(* IEC 61131-3 sources: lasal-git-demo/CPU/LasalDemoProject/Class/_OpenSSL, 1 file *)

(* ---- _OpenSSL.st ---- *)
#include "..\..\Class\_OpenSSL\lsl_openssl.h"

(*!
<Class
	Name               = "_OpenSSL"
	Revision           = "1.9"
	RealtimeTask       = "false"
	CyclicTask         = "false"
	BackgroundTask     = "false"
	Sigmatek           = "true"
	OSInterface        = "true"
	HighPriority       = "false"
	Automatic          = "false"
	UpdateMode         = "Prescan"
	SharedCommandTable = "true"
	Objectsize         = "(284,120)"
	Comment            = "OpenSSL API">
	<Channels>
		<Server Name="ClassSvr" Visualized="false" Initialize="false" WriteProtected="true" Retentive="false"/>
	</Channels>
	<Dependencies>
		<Files>
			<File Path=".\Class\_OpenSSL\DefineCompiler.h" Include="false"/>
			<File Path=".\Class\_OpenSSL\lsl_c_openssl.h" Include="false"/>
			<File Path=".\Class\_OpenSSL\lsl_openssl.h" Include="true"/>
			<File Path=".\Source\code\OsiBaseNew.h" Include="false"/>
			<File Path=".\Source\code\OsiBaseNew.st"/>
		</Files>
	</Dependencies>
	<RevDoku>
		<Owner/>
		<Dokumentation Revision="1.9" Date="2022-09-02" Author="altman" Company="Sigmatek GmbH &amp; Co KG" Description="Fix function parameters for RSA_size and RSA_public_encrypt."/>
		<Dokumentation Revision="1.8" Date="2022-01-21" Author="altman" Company="Sigmatek GmbH &amp; Co KG" Description="The order of the function pointers (LSL_OPENSSL) has been corrected. &#13;&#10;Added new function (BIO_write, PEM_read_bio_RSA_PUBKEY, SHA512, SHA512_Init, SHA512_Update, SHA512_Final)&#13;&#10;Added new define NID_sha512"/>
		<Dokumentation Revision="1.7" Date="2020-05-05" Author="altman" Company="Sigmatek GmbH &amp; Co KG" Description="Added new function (EVP_sha256, SHA256)"/>
		<Dokumentation Revision="1.6" Date="2018-07-18" Author="FucHer" Company="Sigmatek GmbH &amp; Co KG" Description="Added comments for functions and parameters.&#13;&#10;d2i_RSAPrivateKey(): changed data type of parameter &lt;a&gt; from ^Void to ^pVoid.&#13;&#10;ASN1_TIME_set(): changed data type of parameter &lt;tx&gt; from ^DINT to DINT.&#13;&#10;Use dummy functions with a suitable return value."/>
		<Dokumentation Revision="1.5" Date="2018-06-19" Author="altman" Company="Sigmatek GmbH &amp; Co KG" Description="Added new function (X509_get_notBefore, X509_get_notAfter)&#13;&#10;Added new Type (ASN1_TIME)&#13;&#10;"/>
		<Dokumentation Revision="1.4" Date="2018-06-13" Author="altman" Company="Sigmatek GmbH &amp; Co KG" Description="Add new function (X509_cmp_time)&#13;&#10;Correct function parameter and CIL pointer name."/>
		<Dokumentation Revision="1.3" Date="2018-04-10" Author="altman" Company="Sigmatek GmbH &amp; Co KG" Description="Added new functions"/>
		<Dokumentation Revision="1.2" Date="2018-02-07" Author="fucher" Company="Sigmatek GmbH &amp; Co KG" Description="Added dummy functions to prevent fatal &quot;Ldr syntax error&quot; when CIL is not available.&#13;&#10;Removed duplicate entries from aMeths[]. Added missing entries to aMeths[].&#13;&#10;"/>
	</RevDoku>
</Class>
*)
_OpenSSL : CLASS
	TYPE
#pragma pack(push, 1)
	  LSL_OPENSSL : STRUCT
	    udVersion : UDINT;
	    udSize : UDINT;
	    d2i_X509 : pVoid;
	    X509_get_subject_name : pVoid;
	    X509_NAME_get_index_by_NID : pVoid;
	    X509_NAME_get_entry : pVoid;
	    X509_NAME_ENTRY_get_data : pVoid;
	    ASN1_STRING_to_UTF8 : pVoid;
	    OPENSSL_free : pVoid;
	    X509_free : pVoid;
	    SSLeay_version : pVoid;
	    OpenSSL_add_all_algorithms : pVoid;
	    ERR_load_crypto_strings : pVoid;
	    X509_STORE_CTX_get_ex_new_index : pVoid;
	    EVP_cleanup : pVoid;
	    CRYPTO_cleanup_all_ex_data : pVoid;
	    ERR_remove_state : pVoid;
	    ERR_free_strings : pVoid;
	    AES_set_encrypt_key : pVoid;
	    AES_set_decrypt_key : pVoid;
	    AES_cbc_encrypt : pVoid;
	    EVP_sha1 : pVoid;
	    HMAC : pVoid;
	    X509_STORE_free : pVoid;
	    X509_STORE_add_cert : pVoid;
	    SHA1 : pVoid;
	    RAND_bytes : pVoid;
	    RSA_generate_key : pVoid;
	    i2d_RSAPublicKey : pVoid;
	    i2d_RSAPrivateKey : pVoid;
	    d2i_RSAPrivateKey : pVoid;
	    d2i_PublicKey : pVoid;
	    d2i_PrivateKey : pVoid;
	    RSA_free : pVoid;
	    BIO_new_file : pVoid;
	    PEM_read_bio_PrivateKey : pVoid;
	    d2i_PKCS12_bio : pVoid;
	    PKCS12_parse : pVoid;
	    PKCS12_free : pVoid;
	    EVP_PKEY_get1_RSA : pVoid;
	    EVP_PKEY_free : pVoid;
	    BIO_free : pVoid;
	    PEM_write_bio_RSAPrivateKey : pVoid;
	    RSA_size : pVoid;
	    RSA_public_encrypt : pVoid;
	    RSA_private_decrypt : pVoid;
	    RSA_sign : pVoid;
	    ERR_get_error : pVoid;
	    ERR_error_string : pVoid;
	    RSA_verify : pVoid;
	    OBJ_txt2nid : pVoid;
	    X509_NAME_ENTRY_create_by_NID : pVoid;
	    X509_NAME_add_entry : pVoid;
	    X509V3_EXT_conf : pVoid;
	    X509_add_ext : pVoid;
	    X509_EXTENSION_free : pVoid;
	    X509_new : pVoid;
	    X509_set_version : pVoid;
	    X509_get_serialNumber : pVoid;
	    OPENSSL_Realloc : pVoid;
	    ASN1_INTEGER_set : pVoid;
	    X509_set_pubkey : pVoid;
	    X509_NAME_new : pVoid;
	    X509_set_subject_name : pVoid;
	    X509_set_issuer_name : pVoid;
	    X509_gmtime_adj : pVoid;
	    X509V3_set_ctx : pVoid;
	    X509_sign : pVoid;
	    X509_NAME_free : pVoid;
	    i2d_X509_bio : pVoid;
	    d2i_X509_bio : pVoid;
	    PEM_read_bio_X509 : pVoid;
	    X509_get_pubkey : pVoid;
	    OBJ_obj2nid : pVoid;
	    BIO_new : pVoid;
	    i2d_X509 : pVoid;
	    X509_verify : pVoid;
	    X509_STORE_new : pVoid;
	    CRYPTO_add_lock : pVoid;
	    X509_LOOKUP_file : pVoid;
	    X509_LOOKUP_ctrl : pVoid;
	    X509_verify_cert : pVoid;
	    X509_NAME_oneline : pVoid;
	    X509_load_crl_file : pVoid;
	    X509_STORE_CTX_new : pVoid;
	    X509_STORE_CTX_free : pVoid;
	    X509_STORE_CTX_init : pVoid;
	    X509_get_issuer_name : pVoid;
	    X509_LOOKUP_hash_dir : pVoid;
	    X509_STORE_set_flags : pVoid;
	    X509_STORE_add_lookup : pVoid;
	    X509_STORE_set_default_paths : pVoid;
	    X509_STORE_CTX_get_ex_data : pVoid;
	    X509_STORE_CTX_set_ex_data : pVoid;
	    X509_STORE_CTX_get_error : pVoid;
	    X509_STORE_CTX_get_current_cert : pVoid;
	    X509_STORE_CTX_get_error_depth : pVoid;
	    X509_verify_cert_error_string : pVoid;
	    i2d_PublicKey : pVoid;
	    EVP_PKEY_type : pVoid;
	    CRYPTO_realloc : pVoid;
	    BIO_ctrl : pVoid;
	    BIO_s_mem : pVoid;
	    BIO_s_file : pVoid;
	    X509_get_ext : pVoid;
	    EVP_PKEY_cmp : pVoid;
	    EVP_PKEY_new : pVoid;
	    ASN1_TIME_set : pVoid;
	    X509_CRL_sign : pVoid;
	    X509_PUBKEY_get : pVoid;
	    EVP_PKEY_assign : pVoid;
	    X509V3_EXT_print : pVoid;
	    X509_get_ext_by_NID : pVoid;
	    X509_CRL_set_version : pVoid;
	    X509_CRL_add0_revoked : pVoid;
	    X509_CRL_add1_ext_i2d : pVoid;
	    X509_CRL_set_lastUpdate : pVoid;
	    X509_CRL_set_nextUpdate : pVoid;
	    X509_NAME_add_entry_by_txt : pVoid;
	    X509_REVOKED_set_revocationDate : pVoid;
	    X509_CRL_set_issuer_name : pVoid;
	    X509_REVOKED_set_serialNumber : pVoid;
	    X509_NAME_ENTRY_free : pVoid;
	    X509_CRL_new : pVoid;
	    X509_CRL_free : pVoid;
	    ASN1_TIME_free : pVoid;
	    ASN1_INTEGER_new : pVoid;
	    ASN1_INTEGER_free : pVoid;
	    X509_REVOKED_new : pVoid;
	    X509_REVOKED_free : pVoid;
	    PEM_write_bio_X509_CRL : pVoid;
	    X509_cmp_time : pVoid;
	    X509_get_notBefore : pVoid;
	    X509_get_notAfter : pVoid;
	    EVP_sha256 : pVoid;
	    SHA256 : pVoid;
	    BIO_write : pVoid;
	    PEM_read_bio_RSA_PUBKEY : pVoid;
	    SHA512_Init : pVoid;
	    SHA512_Update : pVoid;
	    SHA512_Final : pVoid;
	    SHA512 : pVoid;
	  END_STRUCT;
#pragma pack(pop)
	END_TYPE
  //Servers:
	ClassSvr 	: SvrChCmd_DINT;
  //Clients:
  //Variables:
  //Functions:

	FUNCTION _OpenSSL
		VAR_OUTPUT
			ret_code 	: ConfStates;
		END_VAR;
				//! <Function Comment="Get the version of the OS interface." Name="GetVersion"/>
	FUNCTION VIRTUAL GLOBAL GetVersion
		VAR_OUTPUT
			ret0 	: UDINT;			//! <Variable Comment="&lt;&gt;0: version number of the OS interface&#13;&#10;  =0: error, no OpenSSL interface available." Name="GetVersion.ret0"/>
		END_VAR;
				//! <Function Comment="d2i_X509() attempts to decode &lt;len&gt; bytes at *&lt;in&gt;. If successful a pointer to the X509 structure is returned. If an error occurred, then NULL is returned.&#13;&#10;If &lt;px&gt; is not NULL, then the returned structure is written to *&lt;px&gt;. If *&lt;px&gt; is not NULL, then it is assumed that *&lt;px&gt; contains a valid X509 structure and an attempt is made to reuse it.&#13;&#10;This &quot;reuse&quot; capability is present for historical compatibility but its use is strongly discouraged (see BUGS in www.openssl.org/docs/man1.0.2/crypto/d2i_X509.html).&#13;&#10;&#13;&#10;NOTES&#13;&#10;The letters i and d in i2d_TYPE stand for &quot;internal&quot; (that is, an internal C structure) and &quot;DER&quot; respectively. So i2d_TYPE converts from internal to DER.&#13;&#10;&#13;&#10;If the call is successful *&lt;in&gt; is incremented to the byte following the parsed data.&#13;&#10;&#13;&#10;See also www.openssl.org/docs/man1.0.2/crypto/d2i_X509.html" Name="d2i_X509"/>
	FUNCTION __CDECL VIRTUAL GLOBAL d2i_X509
		VAR_INPUT
			px 	: ^pVoid;			//! <Variable Comment="Pointer to pointer to X509 structure (i.e. **X509).&#13;&#10;If &lt;px&gt; is not NULL, then the returned structure is written to *&lt;px&gt;." Name="d2i_X509.px"/>
			in 	: ^pChar;			//! <Variable Comment="Pointer to pointer to input buffer (i.e. **char)." Name="d2i_X509.in"/>
			len 	: DINT;			//! <Variable Comment="Number of bytes to decode." Name="d2i_X509.len"/>
		END_VAR
		VAR_OUTPUT
			RetAddr (EAX) 	: ^void;			//! <Variable Comment="If successful a pointer to the X509 structure is returned.&#13;&#10;If an error occurred, then NULL is returned. The error code that can be obtained by ERR_get_error()." Name="d2i_X509.RetAddr"/>
		END_VAR;
				//! <Function Comment="X509_get_subject_name() returns the subject name of certificate &lt;a&gt;. The returned value is an internal pointer which MUST NOT be freed.&#13;&#10;&#13;&#10;See also www.openssl.org/docs/man1.1.0/crypto/X509_get_subject_name.html" Name="X509_get_subject_name"/>
	FUNCTION __CDECL VIRTUAL GLOBAL X509_get_subject_name
		VAR_INPUT
			a 	: ^void;			//! <Variable Comment="Pointer to an X509 structure holding certificate &lt;a&gt;." Name="X509_get_subject_name.a"/>
		END_VAR
		VAR_OUTPUT
			RetAddr (EAX) 	: ^void;			//! <Variable Comment="RetAddr is a pointer to an X509_NAME structure.&#13;&#10;This pointer is an internal pointer which MUST NOT be freed." Name="X509_get_subject_name.RetAddr"/>
		END_VAR;
				//! <Function Comment="X509_NAME_get_index_by_NID() retrieves the next index matching &lt;nid&gt; after &lt;lastpos&gt;. &lt;lastpos&gt; should initially be set to -1.&#13;&#10;If there are no more entries -1 is returned. If &lt;nid&gt; is invalid (doesn&apos;t correspond to a valid OID) then -2 is returned.&#13;&#10;&#13;&#10;See also www.openssl.org/docs/man1.0.2/crypto/X509_NAME_get_entry.html" Name="X509_NAME_get_index_by_NID"/>
	FUNCTION __CDECL VIRTUAL GLOBAL X509_NAME_get_index_by_NID
		VAR_INPUT
			name 	: ^void;			//! <Variable Comment="Pointer to X509_NAME structure." Name="X509_NAME_get_index_by_NID.name"/>
			nid 	: DINT;			//! <Variable Comment="NID.&#13;&#10;Applications which could pass invalid NIDs to X509_NAME_get_index_by_NID() should check for the return value of -2." Name="X509_NAME_get_index_by_NID.nid"/>
			lastpos 	: DINT;			//! <Variable Comment="&lt;lastpos&gt; should initially be set to -1" Name="X509_NAME_get_index_by_NID.lastpos"/>
		END_VAR
		VAR_OUTPUT
			RetVal (EAX) 	: DINT;			//! <Variable Comment="Index of the next matching entry or -1 if not found.&#13;&#10;Method can also return -2 if the supplied NID is invalid." Name="X509_NAME_get_index_by_NID.RetVal"/>
		END_VAR;
				//! <Function Comment="X509_NAME_get_entry() retrieves the X509_NAME_ENTRY from &lt;name&gt; corresponding to index &lt;loc&gt;.&#13;&#10;Acceptable values for &lt;loc&gt; run from 0 to (X509_NAME_entry_count(&lt;name&gt;) - 1).&#13;&#10;The value returned is an internal pointer which must not be freed.&#13;&#10;&#13;&#10;See also www.openssl.org/docs/man1.0.2/crypto/X509_NAME_get_entry.html" Name="X509_NAME_get_entry"/>
	FUNCTION __CDECL VIRTUAL GLOBAL X509_NAME_get_entry
		VAR_INPUT
			name 	: ^void;			//! <Variable Comment="Pointer to X509_NAME structure." Name="X509_NAME_get_entry.name"/>
			loc 	: DINT;			//! <Variable Comment="0 to (X509_NAME_entry_count(name) - 1)" Name="X509_NAME_get_entry.loc"/>
		END_VAR
		VAR_OUTPUT
			RetAddr (EAX) 	: ^void;			//! <Variable Comment="Pointer to an X509_NAME_ENTRY structure.&#13;&#10;This is an internal pointer which MUST NOT be freed." Name="X509_NAME_get_entry.RetAddr"/>
		END_VAR;
				//! <Function Comment="X509_NAME_ENTRY_get_data() retrieves the field value of &lt;NeAddr&gt; in an ASN1_STRING structure.&#13;&#10;&#13;&#10;See also www.openssl.org/docs/man1.1.0/crypto/X509_NAME_ENTRY_get_data.html" Name="X509_NAME_ENTRY_get_data"/>
	FUNCTION __CDECL VIRTUAL GLOBAL X509_NAME_ENTRY_get_data
		VAR_INPUT
			NeAddr 	: ^void;			//! <Variable Comment="Pointer to X509_NAME_ENTRY structure." Name="X509_NAME_ENTRY_get_data.NeAddr"/>
		END_VAR
		VAR_OUTPUT
			RetAddr (EAX) 	: ^void;			//! <Variable Comment="Pointer to ASN1_STRING structure." Name="X509_NAME_ENTRY_get_data.RetAddr"/>
		END_VAR;
				//! <Function Comment="ASN1_STRING_to_UTF8() converts the string &lt;in&gt; to UTF8 format, the converted data is allocated in a buffer in *&lt;out&gt;.&#13;&#10;The length of &lt;out&gt; is returned or a negative error code. The buffer *&lt;out&gt; should be freed using OPENSSL_free().&#13;&#10;&#13;&#10;See also www.openssl.org/docs/man1.1.0/crypto/ASN1_STRING_to_UTF8.html" Name="ASN1_STRING_to_UTF8"/>
	FUNCTION __CDECL VIRTUAL GLOBAL ASN1_STRING_to_UTF8
		VAR_INPUT
			out 	: ^pChar;			//! <Variable Comment="Pointer to pointer to output buffer (i.e. **char)." Name="ASN1_STRING_to_UTF8.out"/>
			in 	: ^void;			//! <Variable Comment="Pointer to ASN1_STRING structure." Name="ASN1_STRING_to_UTF8.in"/>
		END_VAR
		VAR_OUTPUT
			RetVal (EAX) 	: DINT;			//! <Variable Comment="The length of &lt;out&gt; or a negative error code." Name="ASN1_STRING_to_UTF8.RetVal"/>
		END_VAR;
				//! <Function Comment="OPENSSL_free() is like the C free() function.&#13;&#10;&#13;&#10;See also www.openssl.org/docs/man1.1.0/crypto/OPENSSL_malloc.html" Name="OPENSSL_free"/>
	FUNCTION __CDECL VIRTUAL GLOBAL OPENSSL_free
		VAR_INPUT
			Addr 	: ^void;			//! <Variable Comment="Void pointer to the buffer that should be freed." Name="OPENSSL_free.Addr"/>
		END_VAR;
				//! <Function Comment="X509_free() frees up the X509 structure &lt;a&gt;.&#13;&#10;&#13;&#10;See also www.openssl.org/docs/man1.0.2/crypto/X509_free.html" Name="X509_free"/>
	FUNCTION __CDECL VIRTUAL GLOBAL X509_free
		VAR_INPUT
			a 	: ^void;			//! <Variable Comment="Pointer to an X509 structure." Name="X509_free.a"/>
		END_VAR;
				//! <Function Comment="SSLeay_version() returns a pointer to a constant string describing the version of the OpenSSL library or giving information about the library build.&#13;&#10;&#13;&#10;See also www.openssl.org/docs/man1.0.2/crypto/SSLeay_version.html" Name="SSLeay_version"/>
	FUNCTION __CDECL VIRTUAL GLOBAL SSLeay_version
		VAR_INPUT
			info_type 	: DINT;			//! <Variable Comment="The following values are supported:&#13;&#10;&#13;&#10;SSLEAY_VERSION&#13;&#10;  The version of the OpenSSL library including the release date.&#13;&#10;SSLEAY_CFLAGS&#13;&#10;  The compiler flags set for the compilation process in the form &quot;compiler: ...&quot; if available or &quot;compiler: information not available&quot; otherwise.&#13;&#10;SSLEAY_BUILT_ON&#13;&#10;  The date of the build process in the form &quot;built on: ...&quot; if available or &quot;built on: date not available&quot; otherwise.&#13;&#10;SSLEAY_PLATFORM&#13;&#10;  The &quot;Configure&quot; target of the library build in the form &quot;platform: ...&quot; if available or &quot;platform: information not available&quot; otherwise.&#13;&#10;SSLEAY_DIR&#13;&#10;  The &quot;OPENSSLDIR&quot; setting of the library build in the form &quot;OPENSSLDIR: &quot;...&quot; if available or &quot;OPENSSLDIR: N/A&quot; otherwise.&#13;&#10;" Name="SSLeay_version.info_type"/>
		END_VAR
		VAR_OUTPUT
			RetAddr (EAX) 	: ^CHAR;			//! <Variable Comment="The following return values can occur:&#13;&#10;&quot;not available&quot;&#13;&#10;  An invalid value for info_type was given.&#13;&#10;Pointer to constant string&#13;&#10;  Textual description.&#13;&#10;" Name="SSLeay_version.RetAddr"/>
		END_VAR;
				//! <Function Comment="OpenSSL keeps an internal table of digest algorithms and ciphers. It uses this table to lookup ciphers via functions such as EVP_get_cipher_byname().&#13;&#10;OpenSSL_add_all_algorithms() adds all algorithms (digests and ciphers) to the table.&#13;&#10;&#13;&#10;See also www.openssl.org/docs/man1.1.0/crypto/OpenSSL_add_all_algorithms.html&#13;&#10;and       https://wiki.openssl.org/index.php/Libcrypto_API" Name="OpenSSL_add_all_algorithms"/>
	FUNCTION __CDECL VIRTUAL GLOBAL OpenSSL_add_all_algorithms;
				//! <Function Comment="ERR_load_crypto_strings() registers the error strings for all libcrypto functions.&#13;&#10;This function should be called before generating textual error messages. However, this is not required when memory usage is an issue.&#13;&#10;&#13;&#10;See also www.openssl.org/docs/man1.0.2/crypto/ERR_load_crypto_strings.html&#13;&#10;and       https://wiki.openssl.org/index.php/Libcrypto_API" Name="ERR_load_crypto_strings"/>
	FUNCTION __CDECL VIRTUAL GLOBAL ERR_load_crypto_strings;
				//! <Function Comment="The X509_STORE_CTX_get_ex_new_index() function is initially called to &quot;register&quot; some new application specific data.&#13;&#10;It takes three optional function pointers which are called when the parent structure (in this case an RSA structure) is initially created, when it is copied and when it is freed up.&#13;&#10;If any or all of these function pointer arguments are not used they should be set to NULL.&#13;&#10;It also takes additional long and pointer parameters which will be passed to the supplied functions new_func(), dup_func() and free_func() but which otherwise have no special meaning.&#13;&#10;&#13;&#10;See also www.openssl.org/docs/man1.0.2/crypto/X509_STORE_CTX_get_ex_new_index.html&#13;&#10;and       www.openssl.org/docs/man1.0.2/crypto/RSA_get_ex_new_index.html" Name="X509_STORE_CTX_get_ex_new_index"/>
	FUNCTION __CDECL VIRTUAL GLOBAL X509_STORE_CTX_get_ex_new_index
		VAR_INPUT
			argl 	: DINT;			//! <Variable Comment="Will be passed to the supplied functions &lt;new_func&gt;, &lt;dup_func&gt;, &lt;free_func&gt;." Name="X509_STORE_CTX_get_ex_new_index.argl"/>
			argp 	: ^void;			//! <Variable Comment="Will be passed to the supplied functions &lt;new_func&gt;, &lt;dup_func&gt;, &lt;free_func&gt;." Name="X509_STORE_CTX_get_ex_new_index.argp"/>
			new_func 	: ^void;			//! <Variable Comment="Optional function pointer CRYPTO_EX_new which is called when the parent structure (in this case an RSA structure) is initially created.&#13;&#10;&#13;&#10;typedef int CRYPTO_EX_new(void *parent, void *ptr, CRYPTO_EX_DATA *ad, int idx, long argl, void *argp);" Name="X509_STORE_CTX_get_ex_new_index.new_func"/>
			dup_func 	: ^void;			//! <Variable Comment="Optional function pointer CRYPTO_EX_dup which is called when the parent structure (in this case an RSA structure) is copied.&#13;&#10;&#13;&#10;typedef int CRYPTO_EX_dup(CRYPTO_EX_DATA *to, CRYPTO_EX_DATA *from, void *from_d, int idx, long argl, void *argp);" Name="X509_STORE_CTX_get_ex_new_index.dup_func"/>
			free_func 	: ^void;			//! <Variable Comment="Optional function pointer CRYPTO_EX_free which is called when the parent structure (in this case an RSA structure) is freed up.&#13;&#10;&#13;&#10;typedef void CRYPTO_EX_free(void *parent, void *ptr, CRYPTO_EX_DATA *ad, int idx, long argl, void *argp);" Name="X509_STORE_CTX_get_ex_new_index.free_func"/>
		END_VAR
		VAR_OUTPUT
			RetVal (EAX) 	: DINT;			//! <Variable Comment="Returns a new index or -1 on failure (note 0 is a valid index value).&#13;&#10;Each successful call will return an index greater than any previously returned." Name="X509_STORE_CTX_get_ex_new_index.RetVal"/>
		END_VAR;
				//! <Function Comment="EVP_cleanup() removes all ciphers and digests from the table used by OpenSSL_add_all_algorithms().&#13;&#10;&#13;&#10;See also www.openssl.org/docs/man1.0.2/crypto/OpenSSL_add_all_algorithms.html&#13;&#10;and       https://wiki.openssl.org/index.php/Libcrypto_API" Name="EVP_cleanup"/>
	FUNCTION __CDECL VIRTUAL GLOBAL EVP_cleanup;
				//! <Function Comment="OpenSSL provides two primary libraries: libssl and libcrypto. The libcrypto library provides the fundamental cryptographic routines used by libssl. &#13;&#10;You can however use libcrypto without using libssl. In order to use libcrypto it must first be initialised.&#13;&#10;Call EVP_cleanup() and CRYPTO_cleanup_all_ex_data() do to the necessary cleanup after using the libcrypto routines.&#13;&#10;&#13;&#10;See also https://wiki.openssl.org/index.php/Libcrypto_API" Name="CRYPTO_cleanup_all_ex_data"/>
	FUNCTION __CDECL VIRTUAL GLOBAL CRYPTO_cleanup_all_ex_data;
				//! <Function Comment="ERR_remove_state() frees the error queue associated with the current thread.&#13;&#10;Since threads in OpenSSL are no longer identified by unsigned long values any argument to this function is ignored.&#13;&#10;&#13;&#10;Since error queue data structures are allocated automatically for new threads, they must be freed when threads are terminated in order to avoid memory leaks.&#13;&#10;&#13;&#10;See also www.openssl.org/docs/man1.0.2/crypto/ERR_remove_state.html" Name="ERR_remove_state"/>
	FUNCTION __CDECL VIRTUAL GLOBAL ERR_remove_state
		VAR_INPUT
			pid 	: UDINT;			//! <Variable Comment="Since threads in OpenSSL are no longer identified by unsigned long values any argument to this function is ignored." Name="ERR_remove_state.pid"/>
		END_VAR;
				//! <Function Comment="ERR_free_strings() frees all previously loaded error strings.&#13;&#10;&#13;&#10;See also www.openssl.org/docs/man1.0.2/crypto/ERR_free_strings.html" Name="ERR_free_strings"/>
	FUNCTION __CDECL VIRTUAL GLOBAL ERR_free_strings;
				//! <Function Comment="AES_set_encrypt_key() configures &lt;key&gt; to encrypt with the &lt;bits&gt;-bit key, &lt;userkey&gt;.&#13;&#10;&#13;&#10;&lt;userkey&gt; contains the actual 128-bit AES key. &lt;key&gt; is a data structure holding a transformed version of the &lt;userkey&gt;, for efficiency.&#13;&#10;&#13;&#10;See also https://boringssl.googlesource.com/boringssl/+/2490/include/openssl/aes.h&#13;&#10;and       www.cs.umd.edu/~jkatz/security/example.c" Name="AES_set_encrypt_key"/>
	FUNCTION __CDECL VIRTUAL GLOBAL AES_set_encrypt_key
		VAR_INPUT
			userkey 	: ^USINT;			//! <Variable Comment="Pointer to actual 128-bit AES key." Name="AES_set_encrypt_key.userkey"/>
			bits 	: DINT;			//! <Variable Comment="Number of bits in &lt;userkey&gt;." Name="AES_set_encrypt_key.bits"/>
			key 	: ^void;			//! <Variable Comment="Pointer to an AES_KEY structure. It holds a transformed version of the &lt;userkey&gt;, for efficiency." Name="AES_set_encrypt_key.key"/>
		END_VAR
		VAR_OUTPUT
			RetVal (EAX) 	: DINT;			//! <Variable Comment="WARNING: unlike other OpenSSL functions, this returns zero on success and a negative number on error." Name="AES_set_encrypt_key.RetVal"/>
		END_VAR;
				//! <Function Comment="AES_set_decrypt_key() configures &lt;key&gt; to decrypt with the &lt;bits&gt;-bit key, &lt;userkey&gt;.&#13;&#10;&#13;&#10;&lt;userkey&gt; contains the actual 128-bit AES key. &lt;key&gt; is a data structure holding a transformed version of the &lt;userkey&gt;, for efficiency.&#13;&#10;&#13;&#10;See also https://boringssl.googlesource.com/boringssl/+/2490/include/openssl/aes.h&#13;&#10;and       www.cs.umd.edu/~jkatz/security/example.c" Name="AES_set_decrypt_key"/>
	FUNCTION __CDECL VIRTUAL GLOBAL AES_set_decrypt_key
		VAR_INPUT
			userkey 	: ^USINT;			//! <Variable Comment="Pointer to actual 128-bit AES key." Name="AES_set_decrypt_key.userkey"/>
			bits 	: DINT;			//! <Variable Comment="Number of bits in &lt;userkey&gt;." Name="AES_set_decrypt_key.bits"/>
			key 	: ^void;			//! <Variable Comment="Pointer to an AES_KEY structure. It holds a transformed version of the &lt;userkey&gt;, for efficiency." Name="AES_set_decrypt_key.key"/>
		END_VAR
		VAR_OUTPUT
			RetVal (EAX) 	: DINT;			//! <Variable Comment="WARNING: unlike other OpenSSL functions, this returns zero on success and a negative number on error." Name="AES_set_decrypt_key.RetVal"/>
		END_VAR;
				//! <Function Comment="Low-level symmetric encryption/decryption using the AES block cipher in CBC mode (cipher-block-chaining).&#13;&#10;&#13;&#10;AES_cbc_encrypt() encrypts (or decrypts, if &lt;enc&gt; == AES_DECRYPT) &lt;len&gt; bytes from &lt;in&gt; to &lt;out&gt;.&#13;&#10;The length &lt;len&gt; must be a multiple of the block size.&#13;&#10;&#13;&#10;The initialization vector is an array of 16 bytes containing random data.&#13;&#10;&#13;&#10;See also https://boringssl.googlesource.com/boringssl/+/2490/include/openssl/aes.h&#13;&#10;and       https://tls.mbed.org/kb/how-to/encrypt-with-aes-cbc" Name="AES_cbc_encrypt"/>
	FUNCTION __CDECL VIRTUAL GLOBAL AES_cbc_encrypt
		VAR_INPUT
			in 	: ^USINT;			//! <Variable Comment="Pointer to input buffer." Name="AES_cbc_encrypt.in"/>
			out 	: ^USINT;			//! <Variable Comment="Pointer to output buffer." Name="AES_cbc_encrypt.out"/>
			len 	: DINT;			//! <Variable Comment="Number of bytes. Must be a multiple of the block size (16 bytes).&#13;&#10;&lt;enc&gt; = AES_ENCRYPT: length of the plaintext.&#13;&#10;&lt;enc&gt; = AES_DECRYPT: length of the ciphertext." Name="AES_cbc_encrypt.len"/>
			key 	: ^void;			//! <Variable Comment="Pointer to an AES_KEY structure." Name="AES_cbc_encrypt.key"/>
			ivec 	: ^USINT;			//! <Variable Comment="Pointer to the initialization vector. The initialization vector contains 16 bytes of random data.&#13;&#10;&lt;ivec&gt; will be incremented." Name="AES_cbc_encrypt.ivec"/>
			enc 	: DINT;			//! <Variable Comment="AES_ENCRYPT or AES_DECRYPT." Name="AES_cbc_encrypt.enc"/>
		END_VAR;
				//! <Function Comment="EVP_sha1(): the SHA-1 algorithm which produces a 160-bit output from a given input.&#13;&#10;SHA-1 (Secure Hash Algorithm 1) is a cryptographic hash function standardized in NIST FIPS 180-4.&#13;&#10;&#13;&#10;EVP_sha1() returns an EVP_MD structure for the SHA1 digest algorithm.&#13;&#10;&#13;&#10;See also www.openssl.org/docs/man1.0.2/crypto/EVP_sha1.html&#13;&#10;and       www.openssl.org/docs/man1.1.1/man3/EVP_sha1.html" Name="EVP_sha1"/>
	FUNCTION __CDECL VIRTUAL GLOBAL EVP_sha1
		VAR_OUTPUT
			RetAddr (EAX) 	: ^void;			//! <Variable Comment="Pointer to an EVP_MD structure that contains the implementation of the symmetric cipher." Name="EVP_sha1.RetAddr"/>
		END_VAR;
				//! <Function Comment="HMAC is a MAC (message authentication code), i.e. a keyed hash function used for message authentication, which is based on a hash function.&#13;&#10;&#13;&#10;HMAC() computes the message authentication code of the &lt;n_val&gt; bytes at &lt;d_addr&gt; using the hash function &lt;evp_md&gt; and the key &lt;key&gt; which is &lt;key_len&gt; bytes long.&#13;&#10;&#13;&#10;It places the result in &lt;md&gt; (which must have space for the output of the hash function, which is no more than EVP_MAX_MD_SIZE bytes).&#13;&#10;If &lt;md&gt; is NULL, the digest is placed in a static array. The size of the output is placed in &lt;md_len&gt;, unless it is NULL.&#13;&#10;&#13;&#10;See also www.openssl.org/docs/man1.0.2/crypto/hmac.html" Name="HMAC"/>
	FUNCTION __CDECL VIRTUAL GLOBAL HMAC
		VAR_INPUT
			evp_md 	: ^void;			//! <Variable Comment="Pointer to a EVP_MD structure containing the hash function." Name="HMAC.evp_md"/>
			key 	: ^void;			//! <Variable Comment="Void pointer to the key." Name="HMAC.key"/>
			key_len 	: DINT;			//! <Variable Comment="Length of &lt;key&gt; in bytes." Name="HMAC.key_len"/>
			d_addr 	: ^USINT;			//! <Variable Comment="Pointer to input buffer." Name="HMAC.d_addr"/>
			n_val 	: DINT;			//! <Variable Comment="Length of the input buffer in bytes." Name="HMAC.n_val"/>
			md 	: ^USINT;			//! <Variable Comment="Pointer to the result buffer (which must have space for the output of the hash function, which is no more than EVP_MAX_MD_SIZE bytes).&#13;&#10;If &lt;md&gt; is NULL, the digest is placed in a static array (WARNING: not thread-safe)." Name="HMAC.md"/>
			md_len 	: ^UDINT;			//! <Variable Comment="Pointer to the size of the output in &lt;md&gt;." Name="HMAC.md_len"/>
		END_VAR
		VAR_OUTPUT
			RetAddr (EAX) 	: ^USINT;			//! <Variable Comment="HMAC() returns a pointer to the message authentication code or NULL if an error occurred." Name="HMAC.RetAddr"/>
		END_VAR;
				//! <Function Comment="X509_STORE_free() frees up a single X509_STORE object.&#13;&#10;&#13;&#10;See also www.openssl.org/docs/man1.1.0/crypto/X509_STORE_free.html" Name="X509_STORE_free"/>
	FUNCTION __CDECL VIRTUAL GLOBAL X509_STORE_free
		VAR_INPUT
			ctx 	: ^void;			//! <Variable Comment="Pointer to the X509_STORE object." Name="X509_STORE_free.ctx"/>
		END_VAR;
				//! <Function Comment="X509_STORE_add_cert() adds a certificate to the X509_STORE&apos;s local storage.&#13;&#10;Untrusted certificates should not be added in this way.&#13;&#10;&#13;&#10;See also www.openssl.org/docs/manmaster/man3/X509_STORE_add_cert.html&#13;&#10;and       http://www.umich.edu/~x509/ssleay/x509_store.html" Name="X509_STORE_add_cert"/>
	FUNCTION __CDECL VIRTUAL GLOBAL X509_STORE_add_cert
		VAR_INPUT
			ctx 	: ^void;			//! <Variable Comment="Pointer to an X509_STORE object." Name="X509_STORE_add_cert.ctx"/>
			x 	: ^void;			//! <Variable Comment="Pointer to an X509 structure containing a certificate." Name="X509_STORE_add_cert.x"/>
		END_VAR
		VAR_OUTPUT
			RetVal (EAX) 	: DINT;			//! <Variable Comment="Returns 1 on success or 0 on failure." Name="X509_STORE_add_cert.RetVal"/>
		END_VAR;
				//! <Function Comment="SHA-1 (Secure Hash Algorithm) is a cryptographic hash function with a 160 bit output.&#13;&#10;&#13;&#10;SHA1() computes the SHA-1 message digest of the &lt;n_val&gt; bytes at &lt;d_addr&gt; and places it in &lt;md&gt; (which must have space for SHA_DIGEST_LENGTH == 20 bytes of output).&#13;&#10;If &lt;md&gt; is NULL, the digest is placed in a static array. Note: setting &lt;md&gt; to NULL is not thread safe.&#13;&#10;&#13;&#10;See also www.openssl.org/docs/man1.0.2/crypto/SHA1.html" Name="SHA1"/>
	FUNCTION __CDECL VIRTUAL GLOBAL SHA1
		VAR_INPUT
			d_addr 	: ^USINT;			//! <Variable Comment="Pointer to input buffer." Name="SHA1.d_addr"/>
			n_val 	: DINT;			//! <Variable Comment="Length of the input buffer in bytes." Name="SHA1.n_val"/>
			md 	: ^USINT;			//! <Variable Comment="Pointer to the SHA-1 message digest buffer (&lt;md&gt; must have space for SHA_DIGEST_LENGTH == 20 bytes of output). &#13;&#10;If &lt;md&gt; is NULL, the digest is placed in a static array (WARNING: not thread-safe)." Name="SHA1.md"/>
		END_VAR
		VAR_OUTPUT
			RetAddr (EAX) 	: ^USINT;			//! <Variable Comment="Returns a pointer to the hash value." Name="SHA1.RetAddr"/>
		END_VAR;
				//! <Function Comment="RAND_bytes() puts &lt;num&gt; cryptographically strong pseudo-random bytes into &lt;buf&gt;.&#13;&#10;An error occurs if the PRNG has not been seeded with enough randomness to ensure an unpredictable byte sequence.&#13;&#10;&#13;&#10;See also www.openssl.org/docs/man1.0.2/crypto/RAND_bytes.html" Name="RAND_bytes"/>
	FUNCTION __CDECL VIRTUAL GLOBAL RAND_bytes
		VAR_INPUT
			buf 	: ^USINT;			//! <Variable Comment="Pointer to &lt;num&gt; cryptographically strong pseudo-random bytes." Name="RAND_bytes.buf"/>
			num 	: DINT;			//! <Variable Comment="Number of bytes in &lt;buf&gt;." Name="RAND_bytes.num"/>
		END_VAR
		VAR_OUTPUT
			RetVal (EAX) 	: DINT;			//! <Variable Comment="RAND_bytes() returns 1 on success, 0 otherwise.&#13;&#10;The error code can be obtained by ERR_get_error().&#13;&#10;The function return -1 if it is not supported by the current RAND method." Name="RAND_bytes.RetVal"/>
		END_VAR;
				//! <Function Comment="RSA_generate_key() generates a key pair and returns a pointer to an RSA structure holding these keys.&#13;&#10;The pseudo-random number generator must be seeded prior to calling RSA_generate_key().&#13;&#10;&#13;&#10;See also www.openssl.org/docs/man1.1.0/crypto/RSA_generate_key.html&#13;&#10;and       www.openssl.org/docs/man1.1.0/crypto/BN_generate_prime.html&#13;&#10;" Name="RSA_generate_key"/>
	FUNCTION __CDECL VIRTUAL GLOBAL RSA_generate_key
		VAR_INPUT
			bits 	: DINT;			//! <Variable Comment="Modulus size in bits. Key sizes with &lt;bits&gt; less than 1024 should be considered insecure." Name="RSA_generate_key.bits"/>
			e 	: UDINT;			//! <Variable Comment="Public exponent. The exponent is an odd number, typically 3, 17 or 65537." Name="RSA_generate_key.e"/>
			callback 	: pVoid;			//! <Variable Comment="Function pointer to old style callback function.&#13;&#10;&#13;&#10;A callback function may be used to provide feedback about the progress of the key generation.&#13;&#10;If &lt;callback&gt; is not NULL, it will be called as follows using the BN_GENCB_call() function described on the BN_generate_prime page.&#13;&#10;&#13;&#10;    While a random prime number is generated, it is called as described in BN_generate_prime.&#13;&#10;&#13;&#10;    When the n-th randomly generated prime is rejected as not suitable for the key, BN_GENCB_call(callback, 2, n) is called.&#13;&#10;&#13;&#10;    When a random p has been found with p-1 relatively prime to e, it is called as BN_GENCB_call(callback, 3, 0).&#13;&#10;&#13;&#10;The process is then repeated for prime q with BN_GENCB_call(callback, 3, 1)." Name="RSA_generate_key.callback"/>
			cb_arg 	: ^void;			//! <Variable Comment="Will be passed to the callback function:  void (*callback)(int, int, void *cb_arg)." Name="RSA_generate_key.cb_arg"/>
		END_VAR
		VAR_OUTPUT
			RetAddr (EAX) 	: ^UDINT;			//! <Variable Comment="Returns a pointer to an RSA structure holding the generated key pair on success or NULL on error." Name="RSA_generate_key.RetAddr"/>
		END_VAR;
				//! <Function Comment="i2d_RSAPublicKey() converts a PKCS#1 RSAPublicKey structure into DER format.&#13;&#10;The usage of this function is similar to the i2d_X509() described in the d2i_X509 manual page.&#13;&#10;&#13;&#10;NOTES&#13;&#10;The RSA structure passed to the public key encoding function should have all the PKCS#1 public key components present.&#13;&#10;&#13;&#10;The encoded data is in binary form and may contain embedded zeroes. Functions such as strlen() will not return the correct length of the encoded structure.&#13;&#10;&#13;&#10;See also www.openssl.org/docs/man1.0.2/crypto/i2d_RSAPublicKey.html&#13;&#10;and       www.openssl.org/docs/manmaster/man3/i2d_RSA_PUBKEY.html" Name="i2d_RSAPublicKey"/>
	FUNCTION __CDECL VIRTUAL GLOBAL i2d_RSAPublicKey
		VAR_INPUT
			a 	: ^void;			//! <Variable Comment="Pointer to a PKCS#1 RSA public key structure." Name="i2d_RSAPublicKey.a"/>
			pp 	: ^pChar;			//! <Variable Comment="Pointer to pointer to output buffer (i.e. **char).&#13;&#10;If &lt;pp&gt; is not NULL, the DER encoded data is written to the buffer at *&lt;pp&gt;, and *&lt;pp&gt; is incremented to point after the data just written.&#13;&#10;If *&lt;pp&gt; is NULL memory will be allocated for a buffer and the encoded data written to it. In this case *&lt;pp&gt; is not incremented and it points to the start of the data just written." Name="i2d_RSAPublicKey.pp"/>
		END_VAR
		VAR_OUTPUT
			RetVal (EAX) 	: DINT;			//! <Variable Comment="Returns the number of bytes successfully encoded or a negative value if an error occurs." Name="i2d_RSAPublicKey.RetVal"/>
		END_VAR;
				//! <Function Comment="i2d_RSAPrivateKey() converts a PKCS#1 RSAPrivateKey structure into DER format.&#13;&#10;The usage of this function is similar to the i2d_X509() described in the d2i_X509 manual page.&#13;&#10;&#13;&#10;NOTES&#13;&#10;The RSA structure passed to the private key encoding functions should have all the PKCS#1 private key components present.&#13;&#10;&#13;&#10;The encoded data is in binary form and may contain embedded zeroes. Functions such as strlen() will not return the correct length of the encoded structure.&#13;&#10;&#13;&#10;The data encoded by the private key functions is unencrypted and therefore offers no private key security.&#13;&#10;&#13;&#10;See also www.openssl.org/docs/man1.0.2/crypto/i2d_RSAPublicKey.html&#13;&#10;and       www.openssl.org/docs/manmaster/man3/i2d_RSA_PUBKEY.html" Name="i2d_RSAPrivateKey"/>
	FUNCTION __CDECL VIRTUAL GLOBAL i2d_RSAPrivateKey
		VAR_INPUT
			a 	: ^void;			//! <Variable Comment="Pointer to a PKCS#1 RSA private key structure." Name="i2d_RSAPrivateKey.a"/>
			pp 	: ^pChar;			//! <Variable Comment="Pointer to pointer to output buffer (i.e. **char).&#13;&#10;If &lt;pp&gt; is not NULL, the DER encoded data is written to the buffer at *&lt;pp&gt;, and *&lt;pp&gt; is incremented to point after the data just written.&#13;&#10;If *&lt;pp&gt; is NULL memory will be allocated for a buffer and the encoded data written to it. In this case *&lt;pp&gt; is not incremented and it points to the start of the data just written." Name="i2d_RSAPrivateKey.pp"/>
		END_VAR
		VAR_OUTPUT
			RetVal (EAX) 	: DINT;			//! <Variable Comment="Returns the number of bytes successfully encoded or a negative value if an error occurs." Name="i2d_RSAPrivateKey.RetVal"/>
		END_VAR;
				//! <Function Comment="d2i_RSAPrivateKey() converts a private key form DER format into a PKCS#1 RSA structure in internal format.&#13;&#10;The usage of this function is similar to the d2i_X509() described in the d2i_X509 manual page.&#13;&#10;&#13;&#10;NOTES&#13;&#10;The RSA structure passed to the private key encoding functions should have all the PKCS#1 private key components present.&#13;&#10;&#13;&#10;The data encoded by the private key functions is unencrypted and therefore offers no private key security.&#13;&#10;&#13;&#10;See also www.openssl.org/docs/man1.0.2/crypto/d2i_RSAPrivateKey.html&#13;&#10;and       www.openssl.org/docs/man1.1.0/crypto/d2i_X509.html" Name="d2i_RSAPrivateKey"/>
	FUNCTION __CDECL VIRTUAL GLOBAL d2i_RSAPrivateKey
		VAR_INPUT
			a 	: ^pVoid;			//! <Variable Comment="Pointer to pointer to RSA output structure (i.e. **RSA) for the private key in internal format.&#13;&#10;&#13;&#10;If successful a pointer to the RSA structure is returned.&#13;&#10;If an error occurred then NULL is returned.&#13;&#10;&#13;&#10;If d2i_RSAPrivateKey() is successful and &lt;a&gt; is not NULL then a pointer to the returned structure is also written to *&lt;a&gt;. &#13;&#10;On a successful return, if *&lt;a&gt; is not NULL then it is assumed that *&lt;a&gt; contains a valid RSA structure and an attempt is made to reuse it. &#13;&#10;This &quot;reuse&quot; capability is present for historical compatibility but its use is strongly discouraged." Name="d2i_RSAPrivateKey.a"/>
			pp 	: ^pChar;			//! <Variable Comment="Pointer to pointer to input buffer (i.e. **char).&#13;&#10;d2i_RSAPrivateKey() attempts to decode &lt;length&gt; bytes at *&lt;pp&gt;. &#13;&#10;If successful *&lt;pp&gt; is incremented to the byte following the parsed data. &#13;&#10; " Name="d2i_RSAPrivateKey.pp"/>
			length 	: DINT;			//! <Variable Comment="Number of bytes in the input buffer *&lt;pp&gt;." Name="d2i_RSAPrivateKey.length"/>
		END_VAR
		VAR_OUTPUT
			RetAddr (EAX) 	: ^UDINT;			//! <Variable Comment="If successful a pointer to the RSA structure is returned.&#13;&#10;If an error occurred then NULL is returned." Name="d2i_RSAPrivateKey.RetAddr"/>
		END_VAR;
				//! <Function Comment="d2i_PublicKey() converts a public key using algorithm &lt;type_val&gt; from DER format into internal format. &#13;&#10;It attempts to use any key specific format or PKCS#8 unencrypted PublicKeyInfo format.&#13;&#10;The &lt;type_val&gt; parameter should be a public key algorithm constant such as EVP_PKEY_RSA. An error occurs if the decoded key does not match &lt;type_val&gt;.&#13;&#10;This function is similar to the d2i_X509() functions; see d2i_X509.&#13;&#10;&#13;&#10;NOTES&#13;&#10;This function uses DER format and unencrypted keys.&#13;&#10;Applications wishing to encrypt or decrypt private keys should use other functions such as d2i_PKC8PrivateKey() instead.&#13;&#10;&#13;&#10;If the *&lt;a&gt; is not NULL when calling d2i_PublicKey() (i.e. an existing structure is being reused) and the key format is PKCS#8 then *&lt;a&gt; will be freed and replaced on a successful call.&#13;&#10;&#13;&#10;See also www.openssl.org/docs/man1.1.0/crypto/d2i_PublicKey.html&#13;&#10;and       www.openssl.org/docs/man1.1.0/crypto/d2i_X509.html" Name="d2i_PublicKey"/>
	FUNCTION __CDECL VIRTUAL GLOBAL d2i_PublicKey
		VAR_INPUT
			type_val 	: DINT;			//! <Variable Comment="Public key algorithm constant (e.g. EVP_PKEY_RSA)." Name="d2i_PublicKey.type_val"/>
			a 	: ^pVoid;			//! <Variable Comment="Pointer to pointer to EVP_PKEY output structure (i.e. **EVP_PKEY) for the public key in internal format.&#13;&#10;&#13;&#10;If successful a pointer to the EVP_PKEY structure is returned.&#13;&#10;If an error occurred then NULL is returned.&#13;&#10;&#13;&#10;If d2i_PublicKey() is successful and &lt;a&gt; is not NULL then a pointer to the returned structure is also written to *&lt;a&gt;. &#13;&#10;On a successful return, if *&lt;a&gt; is not NULL then it is assumed that *&lt;a&gt; contains a valid EVP_PKEY structure and an attempt is made to reuse it. &#13;&#10;This &quot;reuse&quot; capability is present for historical compatibility but its use is strongly discouraged." Name="d2i_PublicKey.a"/>
			pp 	: ^pChar;			//! <Variable Comment="Pointer to pointer to input buffer (i.e. **char).&#13;&#10;d2i_PublicKey() attempts to decode &lt;length&gt; bytes at *&lt;pp&gt;. &#13;&#10;If successful *&lt;pp&gt; is incremented to the byte following the parsed data. &#13;&#10; " Name="d2i_PublicKey.pp"/>
			length 	: DINT;			//! <Variable Comment="Number of bytes in the input buffer *&lt;pp&gt;." Name="d2i_PublicKey.length"/>
		END_VAR
		VAR_OUTPUT
			RetAddr (EAX) 	: ^void;			//! <Variable Comment="d2i_PublicKey() returns a pointer to a valid EVP_KEY structure or NULL if an error occurs.&#13;&#10;The error code can be obtained by calling ERR_get_error()." Name="d2i_PublicKey.RetAddr"/>
		END_VAR;
				//! <Function Comment="d2i_PrivateKey() converts a private key using algorithm &lt;type_val&gt; from DER format into internal format. &#13;&#10;It attempts to use any key specific format or PKCS#8 unencrypted PrivateKeyInfo format.&#13;&#10;The &lt;type_val&gt; parameter should be a public key algorithm constant such as EVP_PKEY_RSA. An error occurs if the decoded key does not match &lt;type_val&gt;.&#13;&#10;&#13;&#10;NOTES&#13;&#10;This function uses DER format and unencrypted keys.&#13;&#10;Applications wishing to encrypt or decrypt private keys should use other functions such as d2i_PKC8PrivateKey() instead.&#13;&#10;&#13;&#10;If the *&lt;a&gt; is not NULL when calling d2i_PrivateKey() (i.e. an existing structure is being reused) and the key format is PKCS#8 then *&lt;a&gt; will be freed and replaced on a successful call.&#13;&#10;&#13;&#10;See also www.openssl.org/docs/man1.1.0/crypto/d2i_PublicKey.html&#13;&#10;and       www.openssl.org/docs/man1.1.0/crypto/d2i_X509.html" Name="d2i_PrivateKey"/>
	FUNCTION __CDECL VIRTUAL GLOBAL d2i_PrivateKey
		VAR_INPUT
			type_val 	: DINT;			//! <Variable Comment="Public key algorithm constant (e.g. EVP_PKEY_RSA).&#13;&#10;" Name="d2i_PrivateKey.type_val"/>
			a 	: ^pVoid;			//! <Variable Comment="Pointer to pointer to EVP_PKEY output structure (i.e. **EVP_PKEY) for the private key in internal format.&#13;&#10;&#13;&#10;If successful a pointer to the EVP_PKEY structure is returned.&#13;&#10;If an error occurred then NULL is returned.&#13;&#10;&#13;&#10;If d2i_PrivateKey() is successful and &lt;a&gt; is not NULL then a pointer to the returned structure is also written to *&lt;a&gt;. &#13;&#10;On a successful return, if *&lt;a&gt; is not NULL then it is assumed that *&lt;a&gt; contains a valid EVP_PKEY structure and an attempt is made to reuse it. &#13;&#10;This &quot;reuse&quot; capability is present for historical compatibility but its use is strongly discouraged." Name="d2i_PrivateKey.a"/>
			pp 	: ^pChar;			//! <Variable Comment="Pointer to pointer to input buffer (i.e. **char).&#13;&#10;d2i_PrivateKey() attempts to decode &lt;length&gt; bytes at *&lt;pp&gt;. &#13;&#10;If successful *&lt;pp&gt; is incremented to the byte following the parsed data. &#13;&#10;" Name="d2i_PrivateKey.pp"/>
			length 	: DINT;			//! <Variable Comment="Number of bytes in the input buffer *&lt;pp&gt;." Name="d2i_PrivateKey.length"/>
		END_VAR
		VAR_OUTPUT
			RetAddr (EAX) 	: ^void;			//! <Variable Comment="d2i_PrivateKey() returns a pointer to a valid EVP_KEY structure or NULL if an error occurs.&#13;&#10;The error code can be obtained by calling ERR_get_error." Name="d2i_PrivateKey.RetAddr"/>
		END_VAR;
				//! <Function Comment="RSA_free() frees the RSA structure and its components. The key is erased before the memory is returned to the system.&#13;&#10;&#13;&#10;See www.openssl.org/docs/man1.0.2/crypto/RSA_free.html" Name="RSA_free"/>
	FUNCTION __CDECL VIRTUAL GLOBAL RSA_free
		VAR_INPUT
			Param 	: ^void;			//! <Variable Comment="Pointer to an RSA structure." Name="RSA_free.Param"/>
		END_VAR;
				//! <Function Comment="BIO_new_file() creates a new file BIO with mode &lt;mode&gt;. The meaning of &lt;mode&gt; is the same as the stdio function fopen().&#13;&#10;E.g. “w+” creates an empty file for both reading and writing. If a file with the same name already exists, its content is erased, and &#13;&#10;the file is considered as a new empty file.&#13;&#10;The BIO_CLOSE flag is set on the returned BIO.&#13;&#10;&#13;&#10;See also www.openssl.org/docs/man1.0.2/crypto/BIO_new_file.html" Name="BIO_new_file"/>
	FUNCTION __CDECL VIRTUAL GLOBAL BIO_new_file
		VAR_INPUT
			filename 	: ^SINT;			//! <Variable Comment="Pointer to the filename." Name="BIO_new_file.filename"/>
			mode 	: ^SINT;			//! <Variable Comment="The meaning of &lt;mode&gt; is the same as the stdio function fopen()." Name="BIO_new_file.mode"/>
		END_VAR
		VAR_OUTPUT
			RetAddr (EAX) 	: ^void;			//! <Variable Comment="Returns a file BIO (i.e. *BIO) or NULL if an error occurred." Name="BIO_new_file.RetAddr"/>
		END_VAR;
				//! <Function Comment="The PEM functions read or write structures in PEM format. In this sense PEM format is simply base64 encoded data surrounded by header lines.&#13;&#10;&#13;&#10;The PrivateKey functions read or write a private key in PEM format using an EVP_PKEY structure.&#13;&#10;The read functions transparently handle traditional and PKCS#8 format encrypted and unencrypted keys.&#13;&#10;&#13;&#10;The PrivateKey read routines can be used in all applications because they handle all formats transparently.&#13;&#10;&#13;&#10;PEM FUNCTION ARGUMENTS&#13;&#10;The PEM read functions all take an argument TYPE **x and return a TYPE * pointer. Where TYPE is whatever structure the function uses. &#13;&#10;If x is NULL, then the parameter is ignored. If x is not NULL but *x is NULL, then the structure returned will be written to *x.&#13;&#10;If neither x nor *x is NULL, then an attempt is made to reuse the structure at *x (but see BUGS and EXAMPLES sections).&#13;&#10;Irrespective of the value of x a pointer to the structure is always returned (or NULL if an error occurred).&#13;&#10;&#13;&#10;If the cb parameters is set to NULL and the u parameter is not NULL, then the u parameter is interpreted as a null terminated string to use as the passphrase.&#13;&#10;For callback details see under cb.&#13;&#10;&#13;&#10;See also www.openssl.org/docs/man1.1.0/crypto/PEM_read_bio_PrivateKey.html" Name="PEM_read_bio_PrivateKey"/>
	FUNCTION __CDECL VIRTUAL GLOBAL PEM_read_bio_PrivateKey
		VAR_INPUT
			bp_addr 	: ^void;			//! <Variable Comment="The &lt;bp_addr&gt; BIO pointer specifies the BIO to read from." Name="PEM_read_bio_PrivateKey.bp_addr"/>
			x 	: ^pVoid;			//! <Variable Comment="A void pointer to a pointer to whatever structure the function uses." Name="PEM_read_bio_PrivateKey.x"/>
			cb 	: ^void;			//! <Variable Comment="NULL or a function pointer to the callback function.&#13;&#10;This is the callback to use when querying for the pass phrase used for encrypted PEM structures (normally only private keys).&#13;&#10;&#13;&#10;The callback routine has the following form:&#13;&#10;&#13;&#10; int cb(char *buf, int size, int rwflag, void *u);&#13;&#10;   buf is the buffer to write the passphrase to.&#13;&#10;   size is the maximum length of the passphrase (i.e. the size of buf).&#13;&#10;   rwflag is a flag which is set to 0 when reading and 1 when writing. A typical routine will ask the user to verify the passphrase (for example by prompting for it twice) if rwflag is 1.&#13;&#10;   The u parameter has the same value as the u parameter passed to the PEM routine. It allows arbitrary data to be passed to the callback by the application (for example a window handle in a GUI application). &#13;&#10;&#13;&#10;The callback must return the number of characters in the passphrase or 0 if an error occurred." Name="PEM_read_bio_PrivateKey.cb"/>
			u 	: ^void;			//! <Variable Comment="If &lt;cb&gt; is set to NULL and &lt;u&gt; is not NULL, then &lt;u&gt; is interpreted as a null terminated string to use as the passphrase.&#13;&#10;If &lt;cb&gt; is not NULL, then &lt;u&gt; is passed to the callback function. See &lt;cb&gt;." Name="PEM_read_bio_PrivateKey.u"/>
		END_VAR
		VAR_OUTPUT
			RetAddr (EAX) 	: ^void;			//! <Variable Comment="Returns either a pointer to the structure read or NULL if an error occurred." Name="PEM_read_bio_PrivateKey.RetAddr"/>
		END_VAR;
				//! <Function Comment="This function converts an OpenSSL object from its ASN.1/DER encoding.&#13;&#10;Unlike the C structures which can have pointers to sub-objects within, the DER is a serialized encoding, suitable for sending over the network, writing to a file, and so on.&#13;&#10;&#13;&#10;d2i_PKCS12_bio() attempts to parse data from BIO &lt;bp_addr&gt;.&#13;&#10;If successful a pointer to the PKCS12 structure is returned.&#13;&#10;If &lt;p12&gt; is not NULL then a pointer to the returned structure is also written to *&lt;p12&gt;. If an error occurred then NULL is returned.&#13;&#10;&#13;&#10;On a successful return, if *&lt;p12&gt; is not NULL then it is assumed that *&lt;p12&gt; contains a valid PKCS12 structure and an attempt is made to reuse it.&#13;&#10;This &quot;reuse&quot; capability is present for historical compatibility but its use is strongly discouraged.&#13;&#10;&#13;&#10;NOTES&#13;&#10;The letters i and d in i2d_TYPE stand for &quot;internal&quot; (that is, an internal C structure) and &quot;DER&quot; respectively. So i2d_TYPE converts from internal to DER.&#13;&#10;The functions can also understand BER forms.&#13;&#10;&#13;&#10;See also www.openssl.org/docs/man1.1.0/crypto/d2i_PKCS12_bio.html" Name="d2i_PKCS12_bio"/>
	FUNCTION __CDECL VIRTUAL GLOBAL d2i_PKCS12_bio
		VAR_INPUT
			bp_addr 	: ^void;			//! <Variable Comment="Pointer to a BIO structure (input in DER format)." Name="d2i_PKCS12_bio.bp_addr"/>
			p12 	: ^pVoid;			//! <Variable Comment="NULL or pointer to pointer to PKCS12 structure (i.e. **PKCS12).&#13;&#10;Output in internal format." Name="d2i_PKCS12_bio.p12"/>
		END_VAR
		VAR_OUTPUT
			RetAddr (EAX) 	: ^void;			//! <Variable Comment="If successful a pointer to the PKCS12 structure is returned.&#13;&#10;If an error occurred then NULL is returned." Name="d2i_PKCS12_bio.RetAddr"/>
		END_VAR;
				//! <Function Comment="PKCS12_parse() parses a PKCS12 structure.&#13;&#10;  &lt;p12&gt; is the PKCS12 structure to parse.&#13;&#10;  &lt;pass&gt; is the passphrase to use.&#13;&#10;&#13;&#10;If successful the private key will be written to *&lt;pkey&gt;, the corresponding certificate to *&lt;cert&gt; and any additional certificates to *&lt;ca&gt;.&#13;&#10;&#13;&#10;NOTES&#13;&#10;The parameters &lt;pkey&gt; and &lt;cert&gt; cannot be NULL.&#13;&#10;&lt;ca&gt; can be &lt;NULL&gt; in which case additional certificates will be discarded.&#13;&#10;*&lt;ca&gt; can also be a valid STACK in which case additional certificates are appended to *&lt;ca&gt;. If *&lt;ca&gt; is NULL a new STACK will be allocated.&#13;&#10;&#13;&#10;The friendlyName and localKeyID attributes (if present) on each certificate will be stored in the alias and keyid attributes of the X509 structure.&#13;&#10;&#13;&#10;The parameter &lt;pass&gt; is interpreted as a string in the UTF-8 encoding. If it is not valid UTF-8, then it is assumed to be ISO8859-1 instead.&#13;&#10;&#13;&#10;In particular, this means that passwords in the locale character set (or code page on Windows) must potentially be converted to UTF-8 before use.&#13;&#10;This may include passwords from local text files, or input from the terminal or command line. Refer to the documentation of UI_OpenSSL(3), for example.&#13;&#10;&#13;&#10;BUGS&#13;&#10;Only a single private key and corresponding certificate is returned by this function. More complex PKCS#12 files with multiple private keys will only return the first match.&#13;&#10;&#13;&#10;Only friendlyName and localKeyID attributes are currently stored in certificates. Other attributes are discarded.&#13;&#10;&#13;&#10;Attributes currently cannot be stored in the private key EVP_PKEY structure.&#13;&#10;&#13;&#10;&#13;&#10;See also www.openssl.org/docs/manmaster/man3/PKCS12_parse.html" Name="PKCS12_parse"/>
	FUNCTION __CDECL VIRTUAL GLOBAL PKCS12_parse
		VAR_INPUT
			p12 	: ^void;			//! <Variable Comment="Pointer to the PKCS12 structure to parse." Name="PKCS12_parse.p12"/>
			pass 	: ^SINT;			//! <Variable Comment="Pointer to the passphrase to use." Name="PKCS12_parse.pass"/>
			pkey 	: ^pVoid;			//! <Variable Comment="Pointer to pointer to an EVP_PKEY structure holding the private key (i.e. **EVP_PKEY)." Name="PKCS12_parse.pkey"/>
			cert 	: ^pVoid;			//! <Variable Comment="Pointer to pointer to a X509 structure holding the corresponding certificate (i.e. **X509)." Name="PKCS12_parse.cert"/>
			ca 	: ^pVoid;			//! <Variable Comment="Pointer to pointer to STACK_OF(X509) holding any additional certificates (i.e. **STACK_OF(X509))." Name="PKCS12_parse.ca"/>
		END_VAR
		VAR_OUTPUT
			RetVal (EAX) 	: DINT;			//! <Variable Comment="PKCS12_parse() returns 1 for success and zero if an error occurred.&#13;&#10;The error can be obtained from ERR_get_error()." Name="PKCS12_parse.RetVal"/>
		END_VAR;
				//! <Function Comment="PKCS12_free() releases the object and all pointers and sub-objects within it.&#13;&#10;&#13;&#10;See also /www.openssl.org/docs/man1.1.0/crypto/PKCS12_free.html" Name="PKCS12_free"/>
	FUNCTION __CDECL VIRTUAL GLOBAL PKCS12_free
		VAR_INPUT
			a 	: ^void;			//! <Variable Comment="Pointer to PKCS12 structure." Name="PKCS12_free.a"/>
		END_VAR;
				//! <Function Comment="EVP_PKEY_get1_RSA() returns the referenced key in &lt;pkey&gt; or NULL if the key is not of the correct type.&#13;&#10;&#13;&#10;NOTES&#13;&#10;In accordance with the OpenSSL naming convention the key obtained from or assigned to the &lt;pkey&gt; must be freed as well as &lt;pkey&gt;.&#13;&#10;&#13;&#10;See also www.openssl.org/docs/man1.0.2/crypto/EVP_PKEY_get1_RSA.html" Name="EVP_PKEY_get1_RSA"/>
	FUNCTION __CDECL VIRTUAL GLOBAL EVP_PKEY_get1_RSA
		VAR_INPUT
			pkey 	: ^void;			//! <Variable Comment="Pointer to an EVP_PKEY structure." Name="EVP_PKEY_get1_RSA.pkey"/>
		END_VAR
		VAR_OUTPUT
			RetAddr (EAX) 	: ^void;			//! <Variable Comment="Returns a pointer to an RSA structure holding the referenced key or NULL if an error occurred." Name="EVP_PKEY_get1_RSA.RetAddr"/>
		END_VAR;
				//! <Function Comment="EVP_PKEY_free() frees up the private key &lt;key&gt;.&#13;&#10;&#13;&#10;See also www.openssl.org/docs/man1.0.2/crypto/EVP_PKEY_free.html" Name="EVP_PKEY_free"/>
	FUNCTION __CDECL VIRTUAL GLOBAL EVP_PKEY_free
		VAR_INPUT
			key 	: ^void;			//! <Variable Comment="Pointer to an EVP_PKEY structure." Name="EVP_PKEY_free.key"/>
		END_VAR;
				//! <Function Comment="BIO_free() frees up a single BIO.&#13;&#10;Calling BIO_free() may also have some effect on the underlying I/O structure, for example it may close the file being referred to under certain circumstances.&#13;&#10;For more details see the individual BIO_METHOD descriptions.&#13;&#10;&#13;&#10;NOTES&#13;&#10;If BIO_free() is called on a BIO chain it will only free one BIO resulting in a memory leak.&#13;&#10;&#13;&#10;See also www.openssl.org/docs/man1.0.2/crypto/BIO_free.html" Name="BIO_free"/>
	FUNCTION __CDECL VIRTUAL GLOBAL BIO_free
		VAR_INPUT
			a 	: ^void;			//! <Variable Comment="Pointer to a BIO structure." Name="BIO_free.a"/>
		END_VAR
		VAR_OUTPUT
			RetVal (EAX) 	: DINT;			//! <Variable Comment="BIO_free() returns 1 for success and 0 for failure." Name="BIO_free.RetVal"/>
		END_VAR;
				//! <Function Comment="The PEM functions read or write structures in PEM format. In this sense PEM format is simply base64 encoded data surrounded by header lines.&#13;&#10;&#13;&#10;The PEM_write_bio_RSAPrivateKey() function processes an RSA private key using an RSA structure. The write routine uses traditional format.&#13;&#10;&#13;&#10;NOTES&#13;&#10;The old PrivateKey write routines are retained for compatibility. New applications should write private keys using the PEM_write_bio_PKCS8PrivateKey() &#13;&#10;or PEM_write_PKCS8PrivateKey() routines because they are more secure (they use an iteration count of 2048 whereas the traditional routines use a count of 1) &#13;&#10;unless compatibility with older versions of OpenSSL is important.&#13;&#10;&#13;&#10;See also www.openssl.org/docs/man1.1.0/crypto/PEM_write_bio_RSAPrivateKey.html" Name="PEM_write_bio_RSAPrivateKey"/>
	FUNCTION __CDECL VIRTUAL GLOBAL PEM_write_bio_RSAPrivateKey
		VAR_INPUT
			bp_addr 	: ^void;			//! <Variable Comment="Pointer to the BIO structure to write to." Name="PEM_write_bio_RSAPrivateKey.bp_addr"/>
			x 	: ^void;			//! <Variable Comment="Pointer to RSA structure holding the private key." Name="PEM_write_bio_RSAPrivateKey.x"/>
			enc 	: ^void;			//! <Variable Comment="Pointer to EVP_CIPHER specifies the encryption algorithm to use. Encryption is done at the PEM level.&#13;&#10;If this parameter is set to NULL then the private key is written in unencrypted form." Name="PEM_write_bio_RSAPrivateKey.enc"/>
			kstr 	: ^USINT;			//! <Variable Comment="If &lt;kstr&gt; is not NULL then &lt;klen&gt; bytes at &lt;kstr&gt; are used as the passphrase and &lt;cb&gt; is ignored." Name="PEM_write_bio_RSAPrivateKey.kstr"/>
			klen 	: DINT;			//! <Variable Comment="If &lt;kstr&gt; is not NULL then &lt;klen&gt; bytes at &lt;kstr&gt; are used as the passphrase and &lt;cb&gt; is ignored." Name="PEM_write_bio_RSAPrivateKey.klen"/>
			cb 	: ^void;			//! <Variable Comment="NULL or a function pointer to the callback function.&#13;&#10;This is the callback to use when querying for the pass phrase used for encrypted PEM structures (normally only private keys).&#13;&#10;&#13;&#10;The callback routine has the following form:&#13;&#10;&#13;&#10; int cb(char *buf, int size, int rwflag, void *u);&#13;&#10;   buf is the buffer to write the passphrase to.&#13;&#10;   size is the maximum length of the passphrase (i.e. the size of buf).&#13;&#10;   rwflag is a flag which is set to 0 when reading and 1 when writing. A typical routine will ask the user to verify the passphrase (for example by prompting for it twice) if rwflag is 1.&#13;&#10;   The u parameter has the same value as the u parameter passed to the PEM routine. It allows arbitrary data to be passed to the callback by the application (for example a window handle in a GUI application). &#13;&#10;&#13;&#10;The callback must return the number of characters in the passphrase or 0 if an error occurred." Name="PEM_write_bio_RSAPrivateKey.cb"/>
			u 	: ^void;			//! <Variable Comment="If &lt;cb&gt; is set to NULL and &lt;u&gt; is not NULL then &lt;u&gt; is interpreted as a null terminated string to use as the passphrase.&#13;&#10;If &lt;cb&gt; is not NULL then &lt;u&gt; is passed to the callback function. See &lt;cb&gt;." Name="PEM_write_bio_RSAPrivateKey.u"/>
		END_VAR
		VAR_OUTPUT
			RetVal (EAX) 	: DINT;			//! <Variable Comment="Returns 1 for success or 0 for failure." Name="PEM_write_bio_RSAPrivateKey.RetVal"/>
		END_VAR;
				//! <Function Comment="This function returns the RSA modulus size in bytes. It can be used to determine how much memory must be allocated for an RSA encrypted value.&#13;&#10;&#13;&#10;rsa-&gt;n must not be NULL.&#13;&#10;&#13;&#10;See also www.openssl.org/docs/man1.0.2/crypto/RSA_size.html" Name="RSA_size"/>
	FUNCTION __CDECL VIRTUAL GLOBAL RSA_size
		VAR_INPUT
			rsa 	: ^void;			//! <Variable Comment="Pointer to RSA structure." Name="RSA_size.rsa"/>
		END_VAR
		VAR_OUTPUT
			RetVal (EAX) 	: DINT;			//! <Variable Comment="The size in bytes." Name="RSA_size.RetVal"/>
		END_VAR;
				//! <Function Comment="The RSA functions implement RSA public key encryption and signatures as defined in PKCS #1 v2.0 [RFC 2437].&#13;&#10;&#13;&#10;RSA_public_encrypt() encrypts the &lt;flen&gt; bytes at &lt;from_addr&gt; (usually a session key) using the public key &lt;rsa&gt; and stores the ciphertext in &lt;to_addr&gt;. &#13;&#10;&lt;to_addr&gt; must point to RSA_size(&lt;rsa&gt;) bytes of memory.&#13;&#10;The random number generator must be seeded prior to calling RSA_public_encrypt().&#13;&#10;&#13;&#10;WARNING&#13;&#10;Decryption failures in the RSA_PKCS1_PADDING mode leak information which can potentially be used to mount a Bleichenbacher padding oracle attack.&#13;&#10;This is an inherent weakness in the PKCS #1 v1.5 padding design. Prefer RSA_PKCS1_OAEP_PADDING.&#13;&#10;&#13;&#10;See also www.openssl.org/docs/man1.0.2/crypto/RSA_public_encrypt.html&#13;&#10;and       www.openssl.org/docs/man1.0.2/crypto/rsa.html" Name="RSA_public_encrypt"/>
	FUNCTION __CDECL VIRTUAL GLOBAL RSA_public_encrypt
		VAR_INPUT
			flen 	: DINT;			//! <Variable Comment="Number of bytes to encrypt.&#13;&#10;&#13;&#10;&lt;flen&gt; must be less than RSA_size(rsa) - 11 for the PKCS #1 v1.5 based padding modes,&#13;&#10;less than RSA_size(rsa) - 41 for RSA_PKCS1_OAEP_PADDING and exactly RSA_size(rsa) for RSA_NO_PADDING." Name="RSA_public_encrypt.flen"/>
			from_addr 	: ^USINT;			//! <Variable Comment="Pointer to the plaintext (data to be encrypted)." Name="RSA_public_encrypt.from_addr"/>
			to_addr 	: ^USINT;			//! <Variable Comment="Pointer to the ciphertext." Name="RSA_public_encrypt.to_addr"/>
			rsa 	: ^void;			//! <Variable Comment="Pointer to an RSA structure holding the public key." Name="RSA_public_encrypt.rsa"/>
			padding 	: DINT;			//! <Variable Comment="&lt;padding&gt; denotes one of the following modes:&#13;&#10;&#13;&#10;RSA_PKCS1_PADDING&#13;&#10;&#13;&#10;    PKCS #1 v1.5 padding. This currently is the most widely used mode.&#13;&#10;RSA_PKCS1_OAEP_PADDING&#13;&#10;&#13;&#10;    EME-OAEP as defined in PKCS #1 v2.0 with SHA-1, MGF1 and an empty encoding parameter. This mode is recommended for all new applications.&#13;&#10;RSA_SSLV23_PADDING&#13;&#10;&#13;&#10;    PKCS #1 v1.5 padding with an SSL-specific modification that denotes that the server is SSL3 capable.&#13;&#10;RSA_NO_PADDING&#13;&#10;&#13;&#10;    Raw RSA encryption. This mode should only be used to implement cryptographically sound padding modes in the application code. Encrypting user data directly with RSA is insecure.&#13;&#10;" Name="RSA_public_encrypt.padding"/>
		END_VAR
		VAR_OUTPUT
			RetVal (EAX) 	: DINT;			//! <Variable Comment="Returns the size of the encrypted data (i.e., RSA_size(rsa)).&#13;&#10;On error, -1 is returned; the error codes can be obtained by ERR_get_error()." Name="RSA_public_encrypt.RetVal"/>
		END_VAR;
				//! <Function Comment="The RSA functions implement RSA public key encryption and signatures as defined in PKCS #1 v2.0 [RFC 2437].&#13;&#10;&#13;&#10;RSA_private_decrypt() decrypts the &lt;flen&gt; bytes at &lt;from_Addr&gt; using the private key &lt;rsa&gt; and stores the plaintext in &lt;to_addr&gt;.&#13;&#10;&lt;to_addr&gt; must point to a memory section large enough to hold the decrypted data (which is smaller than RSA_size(&lt;rsa&gt;)).&#13;&#10;&lt;padding&gt; is the padding mode that was used to encrypt the data.&#13;&#10;&#13;&#10;See also www.openssl.org/docs/man1.0.2/crypto/RSA_public_encrypt.html&#13;&#10;and       www.openssl.org/docs/man1.0.2/crypto/rsa.html" Name="RSA_private_decrypt"/>
	FUNCTION __CDECL VIRTUAL GLOBAL RSA_private_decrypt
		VAR_INPUT
			flen 	: DINT;			//! <Variable Comment="&lt;flen&gt; is RSA_size(&lt;rsa&gt;)." Name="RSA_private_decrypt.flen"/>
			from_Addr 	: ^USINT;			//! <Variable Comment="Pointer to the encrypted ciphertext." Name="RSA_private_decrypt.from_Addr"/>
			to_addr 	: ^USINT;			//! <Variable Comment="Pointer to the decrypted plaintext." Name="RSA_private_decrypt.to_addr"/>
			rsa 	: ^void;			//! <Variable Comment="Pointer to an RSA structure holding the private key." Name="RSA_private_decrypt.rsa"/>
			padding 	: DINT;			//! <Variable Comment="The padding mode that was used to encrypt the data." Name="RSA_private_decrypt.padding"/>
		END_VAR
		VAR_OUTPUT
			RetVal (EAX) 	: DINT;			//! <Variable Comment="RSA_private_decrypt() returns the size of the recovered plaintext.&#13;&#10;On error, -1 is returned; the error codes can be obtained by ERR_get_error()." Name="RSA_private_decrypt.RetVal"/>
		END_VAR;
				//! <Function Comment="RSA_sign() signs the message digest &lt;m_addr&gt; of size &lt;m_len&gt; using the private key &lt;rsa&gt; as specified in PKCS #1 v2.0.&#13;&#10;It stores the signature in &lt;sigret&gt; and the signature size in &lt;siglen&gt;. &lt;sigret&gt; must point to RSA_size(&lt;rsa&gt;) bytes of memory.&#13;&#10;Note that PKCS #1 adds meta-data, placing limits on the size of the key that can be used.&#13;&#10;&#13;&#10;BUGS&#13;&#10;Certain signatures with an improper algorithm identifier are accepted for compatibility with SSLeay 0.4.5 :-)&#13;&#10;&#13;&#10;See also www.openssl.org/docs/man1.0.2/crypto/RSA_sign.html" Name="RSA_sign"/>
	FUNCTION __CDECL VIRTUAL GLOBAL RSA_sign
		VAR_INPUT
			type_val 	: DINT;			//! <Variable Comment="&lt;type_val&gt; denotes the message digest algorithm that was used to generate &lt;m_addr&gt;. It usually is one of NID_sha1, NID_ripemd160 and NID_md5.&#13;&#10;If &lt;type_val&gt; is NID_md5_sha1, an SSL signature (MD5 and SHA1 message digests with PKCS #1 padding and no algorithm identifier) is created." Name="RSA_sign.type_val"/>
			m_addr 	: ^USINT;			//! <Variable Comment="Pointer to the message digest." Name="RSA_sign.m_addr"/>
			m_len 	: DINT;			//! <Variable Comment="Length of the message digest." Name="RSA_sign.m_len"/>
			sigret 	: ^USINT;			//! <Variable Comment="Pointer to the signature." Name="RSA_sign.sigret"/>
			siglen 	: ^UDINT;			//! <Variable Comment="Pointer to the signature size." Name="RSA_sign.siglen"/>
			rsa 	: ^void;			//! <Variable Comment="Pointer to an RSA structure holding the private key as specified in PKCS #1 v2.0." Name="RSA_sign.rsa"/>
		END_VAR
		VAR_OUTPUT
			RetVal (EAX) 	: DINT;			//! <Variable Comment="RSA_sign() returns 1 on success, 0 otherwise." Name="RSA_sign.RetVal"/>
		END_VAR;
				//! <Function Comment="ERR_get_error() returns the earliest error code from the thread&apos;s error queue and removes the entry.&#13;&#10;This function can be called repeatedly until there are no more error codes to return.&#13;&#10;&#13;&#10;See also www.openssl.org/docs/man1.0.2/crypto/ERR_get_error.html" Name="ERR_get_error"/>
	FUNCTION __CDECL VIRTUAL GLOBAL ERR_get_error
		VAR_OUTPUT
			RetVal (EAX) 	: UDINT;			//! <Variable Comment="The error code, or 0 if there is no error in the queue." Name="ERR_get_error.RetVal"/>
		END_VAR;
				//! <Function Comment="ERR_error_string() generates a human-readable string representing the error code &lt;e&gt;, and places it at &lt;buf&gt;.&#13;&#10;&lt;buf&gt; must be at least 120 bytes long. If &lt;buf&gt; is NULL, the error string is placed in a static buffer.&#13;&#10;&#13;&#10;The string will have the following format:&#13;&#10; error:[error code]:[library name]:[function name]:[reason string]&#13;&#10;&#13;&#10;error code is an 8 digit hexadecimal number, library name, function name and reason string are ASCII text.&#13;&#10;&#13;&#10;See also www.openssl.org/docs/man1.0.2/crypto/ERR_error_string.html" Name="ERR_error_string"/>
	FUNCTION __CDECL VIRTUAL GLOBAL ERR_error_string
		VAR_INPUT
			e 	: UDINT;			//! <Variable Comment="Error code." Name="ERR_error_string.e"/>
			buf 	: ^CHAR;			//! <Variable Comment="Pointer to a buffer for the error string.&#13;&#10;The buffer must be at least 120 bytes long.&#13;&#10;If &lt;buf&gt; is NULL, the error string is placed in a static buffer (see RetAddr)." Name="ERR_error_string.buf"/>
		END_VAR
		VAR_OUTPUT
			RetAddr (EAX) 	: ^CHAR;			//! <Variable Comment="ERR_error_string() returns a pointer to a static buffer containing the string if &lt;buf&gt; == NULL, &lt;buf&gt; otherwise." Name="ERR_error_string.RetAddr"/>
		END_VAR;
				//! <Function Comment="RSA_verify() verifies that the signature &lt;sigbuf&gt; of size &lt;siglen&gt; matches a given message digest &lt;m_addr&gt; of size &lt;m_len&gt;.&#13;&#10;&#13;&#10;&lt;rsa&gt; is the signer&apos;s public key.&#13;&#10;&#13;&#10;BUGS&#13;&#10;Certain signatures with an improper algorithm identifier are accepted for compatibility with SSLeay 0.4.5 :-)&#13;&#10;&#13;&#10;See also www.openssl.org/docs/man1.0.2/crypto/RSA_verify.html" Name="RSA_verify"/>
	FUNCTION __CDECL VIRTUAL GLOBAL RSA_verify
		VAR_INPUT
			type_val 	: DINT;			//! <Variable Comment="&lt;type_val&gt; denotes the message digest algorithm that was used to generate the signature." Name="RSA_verify.type_val"/>
			m_addr 	: ^USINT;			//! <Variable Comment="Pointer to the message digest." Name="RSA_verify.m_addr"/>
			m_len 	: UDINT;			//! <Variable Comment="Length of the message digest." Name="RSA_verify.m_len"/>
			sigbuf 	: ^USINT;			//! <Variable Comment="Pointer to the signature." Name="RSA_verify.sigbuf"/>
			siglen 	: UDINT;			//! <Variable Comment="Signature size." Name="RSA_verify.siglen"/>
			rsa 	: ^void;			//! <Variable Comment="Pointer to an RSA structure holding the signer&apos;s public key." Name="RSA_verify.rsa"/>
		END_VAR
		VAR_OUTPUT
			RetVal (EAX) 	: DINT;			//! <Variable Comment="SA_verify() returns 1 on successful verification, 0 otherwise." Name="RSA_verify.RetVal"/>
		END_VAR;
				//! <Function Comment="The ASN1 object utility functions process ASN1_OBJECT structures which are a representation of the ASN1 OBJECT IDENTIFIER (OID) type.&#13;&#10;For convenience, OIDs are usually represented in source code as numeric identifiers, or NIDs.&#13;&#10;OpenSSL has an internal table of OIDs that are generated when the library is built, and their corresponding NIDs are available as defined constants.&#13;&#10;Application code should treat all returned values -- OIDs, NIDs, or names -- as constants.&#13;&#10;&#13;&#10;OBJ_txt2nid() returns NID corresponding to text string &lt;s_addr&gt;. &lt;s_addr&gt; can be a long name, a short name or the numerical representation of an object.&#13;&#10;&#13;&#10;NOTES&#13;&#10;Objects in OpenSSL can have a short name, a long name and a numerical identifier (NID) associated with them.&#13;&#10;A standard set of objects is represented in an internal table. The appropriate values are defined in the header file objects.h.&#13;&#10;&#13;&#10;For example the OID for commonName has the following definitions:&#13;&#10;&#13;&#10; #define SN_commonName                   &quot;CN&quot;&#13;&#10; #define LN_commonName                   &quot;commonName&quot;&#13;&#10; #define NID_commonName                  13&#13;&#10;&#13;&#10;Table objects have certain advantages over other objects: for example their NIDs can be used in a C language switch statement.&#13;&#10;They are also static constant structures which are shared: that is there is only a single constant structure for each table object.&#13;&#10;&#13;&#10;Objects which are not in the table have the NID value NID_undef.&#13;&#10;&#13;&#10;Some objects are used to represent algorithms which do not have a corresponding ASN.1 OBJECT IDENTIFIER encoding (for example no OID currently exists for a particular algorithm).&#13;&#10;As a result they cannot be encoded or decoded as part of ASN.1 structures.&#13;&#10;&#13;&#10;&#13;&#10;See also www.openssl.org/docs/man1.0.2/crypto/OBJ_nid2obj.html" Name="OBJ_txt2nid"/>
	FUNCTION __CDECL VIRTUAL GLOBAL OBJ_txt2nid
		VAR_INPUT
			s_addr 	: ^CHAR;			//! <Variable Comment="Pointer to a text string. The text string can be a long name, a short name or the numerical representation of an object.&#13;&#10;" Name="OBJ_txt2nid.s_addr"/>
		END_VAR
		VAR_OUTPUT
			RetVal (EAX) 	: DINT;			//! <Variable Comment="Returns a NID or NID_undef on error." Name="OBJ_txt2nid.RetVal"/>
		END_VAR;
				//! <Function Comment="X509_NAME_ENTRY_create_by_NID() creates and returns an X509_NAME_ENTRY structure.&#13;&#10;The field name is defined by a NID &lt;nid&gt;.&#13;&#10;The field value to be added is in &lt;bytes&gt; of length &lt;len&gt;. &#13;&#10;If &lt;len&gt; is -1 then the field length is calculated internally using strlen(bytes).&#13;&#10;&#13;&#10;NOTES&#13;&#10;X509_NAME_ENTRY_create_by_NID() is seldom used in practice because X509_NAME_ENTRY structures are &#13;&#10;almost always part of X509_NAME structures and the corresponding X509_NAME functions are typically used &#13;&#10;to create and add new entries in a single operation.&#13;&#10;&#13;&#10;The arguments of this function support similar options to the similarly named one of the corresponding X509_NAME functions such as X509_NAME_add_entry_by_NID(). &#13;&#10;So for example &lt;type_val&gt; can be set to MBSTRING_ASC.&#13;&#10;The use of string types such as MBSTRING_ASC or MBSTRING_UTF8 is strongly recommended for the &lt;type_val&gt; parameter. &#13;&#10;This allows the internal code to correctly determine the type of the field and to apply length checks according to the relevant standards.&#13;&#10;&#13;&#10;BUGS&#13;&#10;&lt;type_val&gt; can still be set to V_ASN1_APP_CHOOSE to use a different algorithm to determine field types. &#13;&#10;Since this form does not understand multicharacter types, performs no length checks and can result in invalid field types its use is strongly discouraged.&#13;&#10;&#13;&#10;See also www.openssl.org/docs/man1.1.0/crypto/X509_NAME_ENTRY_create_by_NID.html&#13;&#10;and       www.openssl.org/docs/man1.0.2/crypto/X509_NAME_add_entry_by_NID.html" Name="X509_NAME_ENTRY_create_by_NID"/>
	FUNCTION __CDECL VIRTUAL GLOBAL X509_NAME_ENTRY_create_by_NID
		VAR_INPUT
			ne_addr 	: ^pVoid;			//! <Variable Comment="Pointer to pointer to X509_NAME_ENTRY structure (i.e. **X509_NAME_ENTRY)." Name="X509_NAME_ENTRY_create_by_NID.ne_addr"/>
			nid 	: DINT;			//! <Variable Comment="NID defining the field name." Name="X509_NAME_ENTRY_create_by_NID.nid"/>
			type_val 	: DINT;			//! <Variable Comment="Type of field.&#13;&#10;Can either be a definition of the type of bytes (such as MBSTRING_ASC) or a standard ASN1 type (such as V_ASN1_IA5STRING).&#13;&#10;&#13;&#10;The use of string types such as MBSTRING_ASC or MBSTRING_UTF8 is strongly recommended for the type parameter. &#13;&#10;This allows the internal code to correctly determine the type of the field and to apply length checks according to the relevant standards. &#13;&#10;This is done using ASN1_STRING_set_by_NID().&#13;&#10;&#13;&#10;If instead an ASN1 type is used no checks are performed and the supplied data in bytes is used directly." Name="X509_NAME_ENTRY_create_by_NID.type_val"/>
			bytes 	: ^USINT;			//! <Variable Comment="Pointer to the field value to be added." Name="X509_NAME_ENTRY_create_by_NID.bytes"/>
			len 	: DINT;			//! <Variable Comment="Length of the field value to be added.&#13;&#10;If &lt;len&gt; is -1 then the field length is calculated internally using strlen(&lt;bytes&gt;)." Name="X509_NAME_ENTRY_create_by_NID.len"/>
		END_VAR
		VAR_OUTPUT
			RetAddr (EAX) 	: ^void;			//! <Variable Comment="Pointer to the new X509_NAME_ENTRY structure." Name="X509_NAME_ENTRY_create_by_NID.RetAddr"/>
		END_VAR;
				//! <Function Comment="X509_NAME_add_entry() adds a copy of X509_NAME_ENTRY structure &lt;ne_addr&gt; to &lt;name&gt;. &#13;&#10;The new entry is added to a position determined by &lt;loc&gt; and &lt;set&gt;. &#13;&#10;Since a copy of &lt;ne_addr&gt; is added &lt;ne_addr&gt; must be freed up after the call.&#13;&#10;&#13;&#10;NOTES&#13;&#10;The &lt;loc&gt; and &lt;set&gt; parameters determine where a new entry should be added. For almost all applications &lt;loc&gt; can be set to -1 and &lt;set&gt; to 0. &#13;&#10;This adds a new entry to the end of name as a single valued RelativeDistinguishedName (RDN).&#13;&#10;&#13;&#10;See also www.openssl.org/docs/man1.0.2/crypto/X509_NAME_add_entry_by_NID.html" Name="X509_NAME_add_entry"/>
	FUNCTION __CDECL VIRTUAL GLOBAL X509_NAME_add_entry
		VAR_INPUT
			name 	: ^void;			//! <Variable Comment="Pointer to X509_NAME structure." Name="X509_NAME_add_entry.name"/>
			ne_addr 	: ^void;			//! <Variable Comment="Pointer to X509_NAME_ENTRY structure holding the data to be copied to &lt;name&gt;." Name="X509_NAME_add_entry.ne_addr"/>
			loc 	: DINT;			//! <Variable Comment="&lt;loc&gt; actually determines the index where the new entry is inserted: if it is -1 it is appended." Name="X509_NAME_add_entry.loc"/>
			set 	: DINT;			//! <Variable Comment="&lt;set&gt; determines how the new type is added. &#13;&#10;If it is zero a new RDN is created.&#13;&#10;&#13;&#10;If &lt;set&gt; is -1 or 1 it is added to the previous or next RDN structure respectively. &#13;&#10;This will then be a multivalued RDN: since multivalue RDNs are very seldom used &lt;set&gt; is almost always set to zero." Name="X509_NAME_add_entry.set"/>
		END_VAR
		VAR_OUTPUT
			RetVal (EAX) 	: DINT;			//! <Variable Comment="Returns 1 for success or 0 if an error occurred." Name="X509_NAME_add_entry.RetVal"/>
		END_VAR;
				//! <Function Comment="This function returns an extension based on a &lt;name&gt; and &lt;value&gt; pair. &#13;&#10;If the&#10; pair will not need to access other sections in a config file (or there is no &#10;config file) then the &lt;conf&gt; parameter can be set to NULL." Name="X509V3_EXT_conf"/>
	FUNCTION __CDECL VIRTUAL GLOBAL X509V3_EXT_conf
		VAR_INPUT
			conf 	: ^void;			//! <Variable Comment="&lt;conf&gt; is the LHASH pointer of the configuration file to use. Can be set to NULL." Name="X509V3_EXT_conf.conf"/>
			ctx 	: ^void;			//! <Variable Comment="Pointer to X509V3_CTX extension context structure. &#13;&#10;&#10;" Name="X509V3_EXT_conf.ctx"/>
			name 	: ^CHAR;			//! <Variable Comment="&lt;name&gt; and &lt;value&gt; pair identifies the extension to be returned." Name="X509V3_EXT_conf.name"/>
			value 	: ^CHAR;			//! <Variable Comment="&lt;name&gt; and &lt;value&gt; pair identifies the extension to be returned." Name="X509V3_EXT_conf.value"/>
		END_VAR
		VAR_OUTPUT
			RetAddr (EAX) 	: ^void;			//! <Variable Comment="Pointer to a X509_EXTENSION structure identified by the &lt;name&gt; and &lt;value&gt; pair." Name="X509V3_EXT_conf.RetAddr"/>
		END_VAR;
				//! <Function Comment="Adds extension &lt;ex&gt; to certificate &lt;x&gt; at position &lt;loc&gt;. If &lt;loc&gt; is -1 the new extension is added to the end. &#13;&#10;The passed extension &lt;ex&gt; is duplicated internally so it must be freed after use.&#13;&#10;&#13;&#10;See also www.openssl.org/docs/man1.1.0/crypto/X509_add_ext.html" Name="X509_add_ext"/>
	FUNCTION __CDECL VIRTUAL GLOBAL X509_add_ext
		VAR_INPUT
			x 	: ^void;			//! <Variable Comment="Pointer to a X509 structure holding a certificate." Name="X509_add_ext.x"/>
			ex 	: ^void;			//! <Variable Comment="Pointer to a X509_EXTENSION structure holding the certificate extension." Name="X509_add_ext.ex"/>
			loc 	: DINT;			//! <Variable Comment="Position within certificate." Name="X509_add_ext.loc"/>
		END_VAR
		VAR_OUTPUT
			RetVal (EAX) 	: DINT;			//! <Variable Comment="Returns &#13;&#10;1 if the operation is successful and &#13;&#10;0 if it fails due to a non-fatal error (extension not found, already exists, cannot be encoded) or &#13;&#10;-1 due to a fatal error such as a memory allocation failure." Name="X509_add_ext.RetVal"/>
		END_VAR;
				//! <Function Comment="X509_EXTENSION_free() releases the object and all pointers and sub-objects within it.&#13;&#10;&#13;&#10;See also /www.openssl.org/docs/man1.1.0/crypto/X509_EXTENSION_free.html" Name="X509_EXTENSION_free"/>
	FUNCTION __CDECL VIRTUAL GLOBAL X509_EXTENSION_free
		VAR_INPUT
			a 	: ^void;			//! <Variable Comment="Pointer to a X509_EXTENSION object." Name="X509_EXTENSION_free.a"/>
		END_VAR;
				//! <Function Comment="X509_new() allocates and initializes a X509 structure.&#13;&#10;&#13;&#10;See also www.openssl.org/docs/man1.0.2/crypto/X509_new.html" Name="X509_new"/>
	FUNCTION __CDECL VIRTUAL GLOBAL X509_new
		VAR_OUTPUT
			RetAddr (EAX) 	: ^void;			//! <Variable Comment="If the allocation fails, X509_new() returns NULL and sets an error code that can be obtained by ERR_get_error(). &#13;&#10;Otherwise it returns a X509 pointer to the newly allocated structure." Name="X509_new.RetAddr"/>
		END_VAR;
				//! <Function Comment="X509_set_version() sets the numerical value of the version field of certificate &lt;x&gt; to &lt;version&gt;.&#13;&#10;&#13;&#10;NOTES&#13;&#10;The version field of certificates, certificate requests and CRLs has a DEFAULT value of v1(0) meaning the field should be omitted for version 1. &#13;&#10;This is handled transparently by these functions.&#13;&#10;&#13;&#10;See also www.openssl.org/docs/man1.1.0/crypto/X509_set_version.html" Name="X509_set_version"/>
	FUNCTION __CDECL VIRTUAL GLOBAL X509_set_version
		VAR_INPUT
			x 	: ^void;			//! <Variable Comment="Pointer to a X509 structure holding the certificate." Name="X509_set_version.x"/>
			version 	: DINT;			//! <Variable Comment="Version number." Name="X509_set_version.version"/>
		END_VAR
		VAR_OUTPUT
			RetVal (EAX) 	: DINT;			//! <Variable Comment="Returns 1 for success and 0 for failure." Name="X509_set_version.RetVal"/>
		END_VAR;
				//! <Function Comment="X509_get_serialNumber() returns the serial number of certificate &lt;x&gt; as an ASN1_INTEGER structure which can be examined or initialised. &#13;&#10;The value returned is an internal pointer which MUST NOT be freed up after the call.&#13;&#10;&#13;&#10;See also www.openssl.org/docs/man1.1.0/crypto/X509_get_serialNumber.html" Name="X509_get_serialNumber"/>
	FUNCTION __CDECL VIRTUAL GLOBAL X509_get_serialNumber
		VAR_INPUT
			x 	: ^void;			//! <Variable Comment="Pointer to a X509 structure holding the certificate." Name="X509_get_serialNumber.x"/>
			RetAddr 	: ^void;			//! <Variable Comment="Returns a pointer to an ASN1_INTEGER structure." Name="X509_get_serialNumber.RetAddr"/>
		END_VAR;
				//! <Function Comment="OpenSSL memory allocation is handled by the OPENSSL_xxx API. &#13;&#10;These are generally macro&apos;s that add the standard C __FILE__ and __LINE__ parameters and call a lower-level CRYPTO_xxx API. &#13;&#10;Some functions do not add those parameters but exist for consistency.&#13;&#10;OPENSSL_malloc(), OPENSSL_realloc(), and OPENSSL_free() are like the C malloc(), realloc(), and free() functions. &#13;&#10;OPENSSL_zalloc() calls memset() to zero the memory before returning.&#13;&#10;&#13;&#10;See also www.openssl.org/docs/man1.1.0/crypto/OPENSSL_realloc.html" Name="OPENSSL_Realloc"/>
	FUNCTION __CDECL VIRTUAL GLOBAL OPENSSL_Realloc
		VAR_INPUT
			addr 	: ^void;			//! <Variable Comment="Pointer to a memory block previously allocated." Name="OPENSSL_Realloc.addr"/>
			num 	: DINT;			//! <Variable Comment="New size for the memory block, in bytes." Name="OPENSSL_Realloc.num"/>
			file 	: ^CHAR;			//! <Variable Comment="The Structured Text __FILE__ parameter." Name="OPENSSL_Realloc.file"/>
			line 	: DINT;			//! <Variable Comment="The Structured Text __LINE__ parameter." Name="OPENSSL_Realloc.line"/>
		END_VAR
		VAR_OUTPUT
			RetAddr (EAX) 	: ^void;			//! <Variable Comment="Returns a void pointer to allocated memory or NULL on error." Name="OPENSSL_Realloc.RetAddr"/>
		END_VAR;
				//! <Function Comment="ASN1_INTEGER_set() sets the value of ASN1_INTEGER &lt;a&gt; to the long value &lt;v&gt;.&#13;&#10;&#13;&#10;NOTES&#13;&#10;In general an ASN1_INTEGER or ASN1_ENUMERATED type can contain an integer of almost arbitrary size and so cannot always be represented by a C int64_t type. &#13;&#10;However in many cases (for example version numbers) they represent small integers which can be more easily manipulated if converted to an appropriate C integer type.&#13;&#10;&#13;&#10;See also www.openssl.org/docs/man1.1.0/crypto/ASN1_INTEGER_set.html" Name="ASN1_INTEGER_set"/>
	FUNCTION __CDECL VIRTUAL GLOBAL ASN1_INTEGER_set
		VAR_INPUT
			a 	: ^void;			//! <Variable Comment="Pointer to a ASN1_INTEGER structure." Name="ASN1_INTEGER_set.a"/>
			v 	: DINT;			//! <Variable Comment="New value for the ASN1_INTEGER &lt;a&gt;." Name="ASN1_INTEGER_set.v"/>
		END_VAR
		VAR_OUTPUT
			RetVal (EAX) 	: DINT;			//! <Variable Comment="Returns 1 for success and 0 for failure. It will only fail if a memory allocation error occurs." Name="ASN1_INTEGER_set.RetVal"/>
		END_VAR;
				//! <Function Comment="X509_set_pubkey() attempts to set the public key for certificate &lt;x&gt; to &lt;pkey&gt;. &#13;&#10;The key &lt;pkey&gt; should be freed up after use.&#13;&#10;&#13;&#10;See also www.openssl.org/docs/man1.1.0/crypto/X509_get_pubkey.html" Name="X509_set_pubkey"/>
	FUNCTION __CDECL VIRTUAL GLOBAL X509_set_pubkey
		VAR_INPUT
			x 	: ^void;			//! <Variable Comment="Pointer to a X509 structure holding the certificate." Name="X509_set_pubkey.x"/>
			pkey 	: ^void;			//! <Variable Comment="Pointer to an EVP_PKEY structure holding the public key for certificate &lt;x&gt;." Name="X509_set_pubkey.pkey"/>
		END_VAR
		VAR_OUTPUT
			RetVal (EAX) 	: DINT;			//! <Variable Comment="Returns 1 for success and 0 for failure." Name="X509_set_pubkey.RetVal"/>
		END_VAR;
				//! <Function Comment="X509_NAME_new() allocates an empty object of type X509_NAME. &#13;&#10;The object returned must be released by calling X509_NAME_free().&#13;&#10;&#13;&#10;See also www.openssl.org/docs/man1.1.0/crypto/X509_NAME_new.html&#13;&#10;and       www.openssl.org/docs/man1.0.2/crypto/x509.html" Name="X509_NAME_new"/>
	FUNCTION __CDECL VIRTUAL GLOBAL X509_NAME_new
		VAR_OUTPUT
			RetAddr (EAX) 	: ^void;			//! <Variable Comment="Returns a X509_NAME pointer to the object or NULL on failure." Name="X509_NAME_new.RetAddr"/>
		END_VAR;
				//! <Function Comment="X509_set_subject_name() sets the subject name of certificate &lt;x&gt; to &lt;name&gt;. &#13;&#10;The name parameter is copied internally and should be freed up when it is no longer needed.&#13;&#10;&#13;&#10;See also www.openssl.org/docs/man1.1.0/crypto/X509_set_subject_name.html" Name="X509_set_subject_name"/>
	FUNCTION __CDECL VIRTUAL GLOBAL X509_set_subject_name
		VAR_INPUT
			x 	: ^void;			//! <Variable Comment="Pointer to a X509 structure holding the certificate." Name="X509_set_subject_name.x"/>
			name 	: ^void;			//! <Variable Comment="Pointer to a X509_NAME structure holding the subject name." Name="X509_set_subject_name.name"/>
		END_VAR
		VAR_OUTPUT
			RetVal (EAX) 	: DINT;			//! <Variable Comment="Returns 1 for success and 0 for failure." Name="X509_set_subject_name.RetVal"/>
		END_VAR;
				//! <Function Comment="X509_set_issuer_name() sets the issuer name of certificate &lt;x&gt; to &lt;name&gt;. &#13;&#10;The name parameter is copied internally and should be freed up when it is no longer needed.&#13;&#10;&#13;&#10;See also www.openssl.org/docs/man1.1.0/crypto/X509_set_subject_name.html" Name="X509_set_issuer_name"/>
	FUNCTION __CDECL VIRTUAL GLOBAL X509_set_issuer_name
		VAR_INPUT
			x 	: ^void;			//! <Variable Comment="Pointer to a X509 structure holding the certificate." Name="X509_set_issuer_name.x"/>
			name 	: ^void;			//! <Variable Comment="Pointer to a X509_NAME structure holding the issuer name." Name="X509_set_issuer_name.name"/>
		END_VAR
		VAR_OUTPUT
			RetVal (EAX) 	: DINT;			//! <Variable Comment="Returns 1 for success and 0 for failure." Name="X509_set_issuer_name.RetVal"/>
		END_VAR;
				//! <Function Comment="Set or get time.&#13;&#10;X509_gmtime_adj() sets the ASN1_UTCTIME structure &lt;s_addr&gt; to the time represented&#10; by &lt;adj&gt;. &#13;&#10;The &lt;adj&gt; value can exceed the number of &#10;seconds in a day. " Name="X509_gmtime_adj"/>
	FUNCTION __CDECL VIRTUAL GLOBAL X509_gmtime_adj
		VAR_INPUT
			s_addr 	: ^void;			//! <Variable Comment="Pointer to ASN1_UTCTIME structure or NULL.&#13;&#10;If &lt;s_addr&gt; is NULL a new ASN1_UTCTIME structure is allocated &#10;and returned." Name="X509_gmtime_adj.s_addr"/>
			adj 	: DINT;			//! <Variable Comment="&lt;adj&gt; contains the time in number of seconds.&#13;&#10;If &lt;adj&gt; is zero the actual time is returned in &lt;RetAddr&gt;." Name="X509_gmtime_adj.adj"/>
		END_VAR
		VAR_OUTPUT
			RetAddr (EAX) 	: ^void;			//! <Variable Comment="Returns a pointer to a ASN1_UTCTIME structure or NULL if an error occurred." Name="X509_gmtime_adj.RetAddr"/>
		END_VAR;
				//! <Function Comment="This function sets up an X509V3_CTX extension context structure with details of the certificate&#10; environment: specifically &#13;&#10;the issuers certificate, &#13;&#10;the subject certificate, &#13;&#10;&#10;the certificate request and the CRL. &#13;&#10;If these are not relevant or not &#10;available then they can be set to NULL. &#13;&#10;The &lt;flags&gt; parameter should be set &#10;to zero.&#13;&#10;&#13;&#10;The purpose of the extension context is to allow the extension code to &#10;access various structures relating to the &quot;environment&quot; of the certificate: &#13;&#10;&#10;for example the issuers certificate or the certificate request.&#13;&#10;" Name="X509V3_set_ctx"/>
	FUNCTION __CDECL VIRTUAL GLOBAL X509V3_set_ctx
		VAR_INPUT
			ctx 	: ^void;			//! <Variable Comment="Pointer to X509V3_CTX extension context structure. &#13;&#10;&#10;&#13;&#10;" Name="X509V3_set_ctx.ctx"/>
			issuer 	: ^void;			//! <Variable Comment="X509 pointer to the issuers certificate. Can be NULL." Name="X509V3_set_ctx.issuer"/>
			subj 	: ^void;			//! <Variable Comment="X509 pointer to the subject certificate. Can be NULL." Name="X509V3_set_ctx.subj"/>
			req 	: ^void;			//! <Variable Comment="X509_REQ pointer to the certificate request. Can be NULL." Name="X509V3_set_ctx.req"/>
			crl 	: ^void;			//! <Variable Comment="X509_CRL pointer to the CRL (Certificate Revocation List). Can be NULL." Name="X509V3_set_ctx.crl"/>
			flags 	: DINT;			//! <Variable Comment="Should be set to zero." Name="X509V3_set_ctx.flags"/>
		END_VAR;
				//! <Function Comment="X509_sign() signs certificate &lt;x&gt; using private key &lt;pkey&gt; and message digest &lt;md&gt; and sets the signature in &lt;x&gt;.&#13;&#10;&#13;&#10;NOTES&#13;&#10;For efficiency reasons and to work around ASN.1 encoding issues the encoding of the signed portion of a certificate, certificate request and CRL is cached internally. &#13;&#10;If the signed portion of the structure is modified the encoding is not always updated meaning a stale version is sometimes used. &#13;&#10;This is not normally a problem because modifying the signed portion will invalidate the signature and signing will always update the encoding.&#13;&#10;&#13;&#10;See also /www.openssl.org/docs/man1.1.0/crypto/X509_sign.html" Name="X509_sign"/>
	FUNCTION __CDECL VIRTUAL GLOBAL X509_sign
		VAR_INPUT
			x 	: ^void;			//! <Variable Comment="Pointer to a X509 structure holding the certificate." Name="X509_sign.x"/>
			pkey 	: ^void;			//! <Variable Comment="Pointer to an EVP_PKEY structure holding the private key for certificate &lt;x&gt;." Name="X509_sign.pkey"/>
			md 	: ^void;			//! <Variable Comment="Pointer to a EVP_MD structure holding the message digest." Name="X509_sign.md"/>
		END_VAR
		VAR_OUTPUT
			RetVal (EAX) 	: DINT;			//! <Variable Comment="Returns the size of the signature in bytes for success and zero for failure." Name="X509_sign.RetVal"/>
		END_VAR;
				//! <Function Comment="X509_NAME_free() releases the object and all pointers and sub-objects within it.&#13;&#10;&#13;&#10;See also www.openssl.org/docs/man1.1.0/crypto/X509_NAME_free.html&#13;&#10;and       www.openssl.org/docs/man1.0.2/crypto/x509.html" Name="X509_NAME_free"/>
	FUNCTION __CDECL VIRTUAL GLOBAL X509_NAME_free
		VAR_INPUT
			a 	: ^void;			//! <Variable Comment="Pointer to the X509_NAME object to be freed." Name="X509_NAME_free.a"/>
		END_VAR;
				//! <Function Comment="i2d_X509_bio() encodes the structure pointed to by &lt;x&gt; into DER format and writes the encoding of the structure &lt;x&gt; to BIO &lt;bp_addr&gt;.&#13;&#10;&#13;&#10;NOTES&#13;&#10;The letters i and d in for example i2d_X509_bio() stand for &quot;internal&quot; (that is an internal C structure) and &quot;DER&quot;. &#13;&#10;So i2d_X509 converts from internal to DER. &#13;&#10;&#13;&#10;The functions can also understand BER forms.&#13;&#10;&#13;&#10;The actual X509 structure passed to i2d_X509_bio() must be a valid populated X509 structure. &#13;&#10;It can not simply be fed with an empty structure such as that returned by X509_new().&#13;&#10;&#13;&#10;The encoded data is in binary form and may contain embedded zeroes. Therefore any FILE pointers or BIOs should be opened in binary mode. &#13;&#10;Functions such as strlen() will not return the correct length of the encoded structure.&#13;&#10;&#13;&#10;See also www.openssl.org/docs/man1.0.2/crypto/d2i_X509_fp.html" Name="i2d_X509_bio"/>
	FUNCTION __CDECL VIRTUAL GLOBAL i2d_X509_bio
		VAR_INPUT
			bp_addr 	: ^void;			//! <Variable Comment="Pointer to a BIO structure (output in DER format)." Name="i2d_X509_bio.bp_addr"/>
			x 	: ^void;			//! <Variable Comment="Pointer to a X509 structure holding the certificate.&#13;&#10;Input in internal format." Name="i2d_X509_bio.x"/>
		END_VAR
		VAR_OUTPUT
			RetVal (EAX) 	: DINT;			//! <Variable Comment="Returns 1 for success and 0 for failure." Name="i2d_X509_bio.RetVal"/>
		END_VAR;
				//! <Function Comment="d2i_X509_bio() attempts to parse data from BIO &lt;bp_addr&gt;. &#13;&#10;If successful a pointer to the X509 structure is returned. If an error occurred then NULL is returned. &#13;&#10;If &lt;x&gt; is not NULL then the returned structure is written to *&lt;x&gt;. &#13;&#10;If *&lt;x&gt; is not NULL then it is assumed that *&lt;x&gt; contains a valid X509 structure and an attempt is made to reuse it. &#13;&#10;&#13;&#10;See also /www.openssl.org/docs/man1.0.2/crypto/d2i_X509_fp.html" Name="d2i_X509_bio"/>
	FUNCTION __CDECL VIRTUAL GLOBAL d2i_X509_bio
		VAR_INPUT
			bp_addr 	: ^void;			//! <Variable Comment="Pointer to a BIO structure (input in DER format)." Name="d2i_X509_bio.bp_addr"/>
			x 	: ^pVoid;			//! <Variable Comment="NULL or pointer to a pointer to a X509 structure holding the certificate.&#13;&#10;Output in internal format." Name="d2i_X509_bio.x"/>
		END_VAR
		VAR_OUTPUT
			RetAddr (EAX) 	: ^void;			//! <Variable Comment="If successful a pointer to the X509 structure is returned.&#13;&#10;If an error occurred then NULL is returned." Name="d2i_X509_bio.RetAddr"/>
		END_VAR;
				//! <Function Comment="The PEM functions read or write structures in PEM format. In this sense PEM format is simply base64 encoded data surrounded by header lines.&#13;&#10;&#13;&#10;PEM_read_bio_X509() reads a certificate in PEM format from the BIO &lt;bp_addr&gt; and returns a pointer to the certificate in internal format.&#13;&#10;&#13;&#10;See also www.openssl.org/docs/man1.0.2/crypto/PEM_read_bio_X509.html" Name="PEM_read_bio_X509"/>
	FUNCTION __CDECL VIRTUAL GLOBAL PEM_read_bio_X509
		VAR_INPUT
			bp_addr 	: ^void;			//! <Variable Comment="Pointer to a BIO structure specifying the BIO to read from." Name="PEM_read_bio_X509.bp_addr"/>
			x 	: ^pVoid;			//! <Variable Comment="Pointer to pointer to a X509 structure.&#13;&#10;&#13;&#10;If &lt;x&gt; is NULL, then the parameter is ignored. If &lt;x&gt; is not NULL but *&lt;x&gt; is NULL, then the structure returned will be written to *&lt;x&gt;. &#13;&#10;If neither &lt;x&gt; nor *&lt;x&gt; is NULL, then an attempt is made to reuse the structure at *&lt;x&gt; (but see BUGS and EXAMPLES sections). &#13;&#10;&#13;&#10;Irrespective of the value of &lt;x&gt; a pointer to the structure is always returned (or NULL if an error occurred)." Name="PEM_read_bio_X509.x"/>
			cb 	: ^void;			//! <Variable Comment="NULL or a function pointer to the callback function.&#13;&#10;This is the callback to use when querying for the pass phrase used for encrypted PEM structures (normally only private keys).&#13;&#10;&#13;&#10;The callback routine has the following form:&#13;&#10;&#13;&#10; int cb(char *buf, int size, int rwflag, void *u);&#13;&#10;   buf is the buffer to write the passphrase to.&#13;&#10;   size is the maximum length of the passphrase (i.e. the size of buf).&#13;&#10;   rwflag is a flag which is set to 0 when reading and 1 when writing. A typical routine will ask the user to verify the passphrase (for example by prompting for it twice) if rwflag is 1.&#13;&#10;   The u parameter has the same value as the u parameter passed to the PEM routine. It allows arbitrary data to be passed to the callback by the application (for example a window handle in a GUI application). &#13;&#10;&#13;&#10;The callback must return the number of characters in the passphrase or 0 if an error occurred." Name="PEM_read_bio_X509.cb"/>
			u 	: ^void;			//! <Variable Comment="If &lt;cb&gt; is set to NULL and &lt;u&gt; is not NULL, then &lt;u&gt; is interpreted as a null terminated string to use as the passphrase.&#13;&#10;If &lt;cb&gt; is not NULL, then &lt;u&gt; is passed to the callback function. See &lt;cb&gt;." Name="PEM_read_bio_X509.u"/>
		END_VAR
		VAR_OUTPUT
			RetAddr (EAX) 	: ^void;			//! <Variable Comment="Pointer to a X509 structure or NULL if an error occurred." Name="PEM_read_bio_X509.RetAddr"/>
		END_VAR;
				//! <Function Comment="X509_get_pubkey() attempts to decode the public key for certificate &lt;x&gt;. &#13;&#10;If successful it returns the public key as an EVP_PKEY pointer with its reference count incremented: this means the returned key must be freed up after use.&#13;&#10;&#13;&#10;See also www.openssl.org/docs/man1.1.0/crypto/X509_REQ_set_pubkey.html" Name="X509_get_pubkey"/>
	FUNCTION __CDECL VIRTUAL GLOBAL X509_get_pubkey
		VAR_INPUT
			x 	: ^void;			//! <Variable Comment="Pointer to a X509 structure holding a certificate." Name="X509_get_pubkey.x"/>
		END_VAR
		VAR_OUTPUT
			RetAddr (EAX) 	: ^void;			//! <Variable Comment="Returns the public key as an EVP_PKEY pointer or NULL if an error occurred." Name="X509_get_pubkey.RetAddr"/>
		END_VAR;
				//! <Function Comment="OBJ_obj2nid() returns the corresponding NID for the object &lt;o&gt; or NID_undef if an error occurred.&#13;&#10;&#13;&#10;See also www.openssl.org/docs/man1.0.2/crypto/OBJ_obj2nid.html" Name="OBJ_obj2nid"/>
	FUNCTION __CDECL VIRTUAL GLOBAL OBJ_obj2nid
		VAR_INPUT
			o 	: ^void;			//! <Variable Comment="Pointer to an object of type ASN1_OBJECT." Name="OBJ_obj2nid.o"/>
		END_VAR
		VAR_OUTPUT
			RetVal (EAX) 	: DINT;			//! <Variable Comment="NID or NID_undef if an error occurred." Name="OBJ_obj2nid.RetVal"/>
		END_VAR;
				//! <Function Comment="The BIO_new() function returns a new BIO using method &lt;t&gt;.&#13;&#10;&#13;&#10;See also www.openssl.org/docs/man1.0.2/crypto/BIO_new.html" Name="BIO_new"/>
	FUNCTION __CDECL VIRTUAL GLOBAL BIO_new
		VAR_INPUT
			t 	: ^void;			//! <Variable Comment="Pointer to BIO_METHOD structure." Name="BIO_new.t"/>
		END_VAR
		VAR_OUTPUT
			RetAddr (EAX) 	: ^void;			//! <Variable Comment="Returns a pointer to the newly created BIO or NULL if the call fails." Name="BIO_new.RetAddr"/>
		END_VAR;
				//! <Function Comment="Encodes the structure pointed to by &lt;x&gt; into DER format. &#13;&#10;If &lt;out&gt; is not NULL it writes the DER encoded data to the buffer at *&lt;out&gt;, and increments &lt;out&gt; to point after the data just written.&#13;&#10;&#13;&#10;See also www.openssl.org/docs/man1.1.0/crypto/i2d_X509.html" Name="i2d_X509"/>
	FUNCTION __CDECL VIRTUAL GLOBAL i2d_X509
		VAR_INPUT
			x 	: ^void;			//! <Variable Comment="Pointer to a X509 structure holding a certificate." Name="i2d_X509.x"/>
			out 	: ^pVoid;			//! <Variable Comment="Pointer to pointer to output buffer (i.e. **unsigned char)." Name="i2d_X509.out"/>
		END_VAR
		VAR_OUTPUT
			RetVal (EAX) 	: DINT;			//! <Variable Comment="Returns the length of the encoded data or a negative value if an error occurred." Name="i2d_X509.RetVal"/>
		END_VAR;
				//! <Function Comment="Verifies the signature of certificate &lt;a&gt; using public key &lt;rx&gt;. Only the signature is checked: no other checks (such as certificate chain validity) are performed.&#13;&#10;&#13;&#10;See also www.openssl.org/docs/man1.1.0/crypto/X509_verify.html" Name="X509_verify"/>
	FUNCTION __CDECL VIRTUAL GLOBAL X509_verify
		VAR_INPUT
			a 	: ^void;			//! <Variable Comment="Pointer to a X509 structure holding a certificate." Name="X509_verify.a"/>
			rx 	: ^void;			//! <Variable Comment="Pointer to EVP_PKEY structure holding the public key." Name="X509_verify.rx"/>
		END_VAR
		VAR_OUTPUT
			Retval (EAX) 	: DINT;			//! <Variable Comment="Returns 1 if the signature is valid and 0 if the signature check fails. &#13;&#10;If the signature could not be checked at all because it was invalid or some other error occurred then -1 is returned." Name="X509_verify.Retval"/>
		END_VAR;
				//! <Function Comment="X509_STORE_new() returns a newly created X509_STORE or NULL if the call fails.&#13;&#10;&#13;&#10;See also www.openssl.org/docs/man1.1.0/crypto/X509_STORE_new.html" Name="X509_STORE_new"/>
	FUNCTION __CDECL VIRTUAL GLOBAL X509_STORE_new
		VAR_OUTPUT
			RetAddr (EAX) 	: ^void;			//! <Variable Comment="Pointer to X509_STORE or NULL if the call fails." Name="X509_STORE_new.RetAddr"/>
		END_VAR;
